(* IEC 61131-3 sources: daoli-st-library/DL_Process (part 66) *)

(* ---- FB_DL_InertPurgeSeq.st ---- *)
(*==============================================================================
 * 组件名称 (Component)  : FB_DL_InertPurgeSeq
 * 溯源说明 (Provenance): 道莅 clean-room 防御性实现（IEC 61131-3 纯净实现，闭源文档仅借语义，零代码行）
 * 所属子库 (Sublibrary) : DL_Process / Sequence
 * 当前版本 (Version)    : 1.0.0
 * 兼容性   (Platform)   : CODESYS 3.5 / TwinCAT 3 / 汇川 InoProShop / 施耐德
 *                         Machine Expert；纯 IEC 61131-3（第 3 版），仅用
 *                         Standard.library 的 TON / TIME_TO_DINT / DINT_TO_TIME
 * 组件分类 (Category)   : 功能块（FUNCTION_BLOCK）· 氮气置换顺控
 * 功能一句话 (Summary)  : 抽真空 → 充氮 → 保压取样 三相同循环置换，氧含量达目标
 *                         即放行，循环耗尽未达标则锁定失败，中止任意拍立即停。
 *
 * 本件存在的意义 (Why this unit exists)
 *   可燃溶剂场合点火/投料前的氮气置换是强制步骤，也是审核最容易被问的
 *   一条。它的逻辑不难，但「相转出必须断输入」这一点几乎每份手写代码都会
 *   踩：三相共用一只 TON，抽真空相残留的 ET 会让充氮相提前结束，或者
 *   保压相一进就走。本件把每相各一只 TON、相转出断输入一拍写成结构约束
 *   （R40 家族第三次事故的共同形态就在这一格）。
 *
 * 单循环定义 (One cycle)
 *   eEvacuate   : 抽真空阀开，tEvac 时间到**且**真空达 fVacOk → 进充氮
 *   eFillN2     : 充氮阀开，tFill 时间到 → 进保压取样
 *   eHoldVerify : 全阀关（保持压力），tHold 后读取氧含量
 *                 ≤ fO2Target → eComplete（信息 01DF）
 *                 否则循环数 +1：未达 uMaxCycles → eCycleDone → 回抽真空（信息 01DE）
 *                 已达 uMaxCycles → eFailed（故障 0313）
 *
 * 中止语义（三件顺控件共用同一段口径）
 *   bAbort **任意拍**生效：先清全部执行输出（三相阀），再回 eIdle；
 *   **不排队、不回退重来、不自动续跑**——中止是人的决定，重启必须由新的
 *   bStart 重新开始。原因：自动续跑会让操作工以为按了一次中止就断电了，
 *   实际设备又自己动起来，这是顺控件最危险的一类行为（R34 家族）。
 *
 * 边界安全 (Boundary)
 *   ① fO2Target <= 0、uMaxCycles = 0 或任一 TIME = 0 → 故障 0311、回 eIdle；
 *   ② bO2SensorOk = FALSE → 故障 0312、**禁止放行**（bDone 恒 FALSE）、三阀全关；
 *      氧分析仪坏掉时置换结果无从判断，继续循环只是白烧氮气；
 *   ③ 循环耗尽未达标 → bFailed := TRUE + 故障 0313；
 *   ④ 抽真空相 tEvac 到而真空未达 → 重新计时继续抽，连续 DL_EVAC_RETRY 次仍未达
 *      → 按「置换无法建立」处理，复用 0313（R90 不加码，理由见头注释）；
 *   ⑤ 三相各一只 TON，相转出以「断输入一拍」标志重启，绝不跨相复用实例；
 *   ⑥ 三阀输出互斥，段 1 先全清、段 7 按状态最多置一路（R72）；
 *   ⑦ CASE 落 ELSE 置 0313 并回 eIdle（兜底复用，R90）；
 *   ⑧ 放空阀编排约定：仅在 eComplete（置换合格）后打开以便泄压放行；
 *      eFailed 与其它相一律关闭——置换失败时保持惰化封闭，交人工处置。
 *
 * 引脚补全声明 (Pin completion)
 *   规格正文要求「真空达 fVacOk」判据，但引脚表未列真空度实测，故补
 *   fVacMeas : REAL [kPa g]。缺此引脚则「抽真空到位」无从判断，只能退化成
 *   纯定时，与本件语义不符。
 *
 * 错误码    : 16#0005_01DE 单循环未达标，进入下一循环——信息级
 *             16#0005_01DF 取样窗内氧含量已达目标——信息级，放行前置条件满足
 *             16#0005_0311 置换参数非法（目标/循环数/时长）——故障级，回 eIdle
 *             16#0005_0312 氧分析仪无效，禁止放行——故障级，三阀全关
 *             16#0005_0313 置换循环耗尽未达标（含状态机兜底与真空建立失败复用，R90）——故障级
 * 码位总账  : 16#0005_01DE 用 / 16#0005_01DF 用 ｜ 16#0005_0311 用 / 16#0005_0312 用 / 16#0005_0313 用
 * 状态机    : E_DL_PurgeState（eIdle / eEvacuate / eFillN2 / eHoldVerify / eCycleDone /
 *             eComplete / eFailed / eFault），CASE 含 ELSE 兜底，ELSE 置 16#0005_0313 并回 eIdle
 * 采样约定  : 每任务周期调用一次；各相时长由引脚给定，不读系统时钟
 * 依赖说明  : 只做组合编排，不复制低层算法；无 DL_ 子库调用
 * 验收向量  : V1 启动 → 抽真空 60 s 且真空 −85 kPa（< −80）→ 充氮 60 s → 保压 30 s
 *               读到 O2 1.2 %（≤ 2.0）→ eComplete，bDone = TRUE，eErr = 01DF
 *             V2 保压后 O2 3.5 %（> 2.0）、uMaxCycles = 3 → uCycleDone = 1，eErr = 01DE，
 *                回抽真空继续（循环主向量）
 *             V3 V2 连续三次未达标 → eFailed，bFailed = TRUE，eErr = 0313（耗尽主向量）
 *             V4 抽真空相 bAbort = TRUE → 三阀同拍全 FALSE，回 eIdle，不续跑（中止主向量）
 *             V5 bO2SensorOk = FALSE → eFault，三阀全关，bDone 恒 FALSE，eErr = 0312
 *             V6 uMaxCycles = 0 → eFault，eErr = 0311，回 eIdle
 *             V7 抽真空 3 次定时到但真空只有 −50 kPa → eFailed，eErr = 0313（真空建立失败复用）
 *             V8 eComplete 且 bStart 仍为 TRUE → 保持 eComplete（不放行丢失）；bStart 落 → eIdle
 * 红线自检  : 全局变量声明零使用 / 外部变量访问零使用 / 物理地址零使用 ｜ 纯 IEC 61131-3 ｜ 无除法
 *             浮点只用大小比较 ｜ 无循环 ｜ 全变量双语同行注释 ｜ ENUM + CASE 含 ELSE
 *             ｜ 三只 TON 在主体前部无条件刷新且各相各一只 ｜ 单拍标志全部预清零
 *             ｜ 阈值常量化，无魔法数
 * 修订历史  : 2026-11-16  v1.0.0  首版入库（R22 · 批 3 · 批处理顺控）
 *============================================================================*)

(*-----------------------------------------------------------------------------
 * 枚举: E_DL_PurgeState（归属本功能块，同文件发布，全库唯一定义）
 * 含义: 氮气置换顺控相位，每个成员在 CASE 中有且仅有一个标签。
 *-----------------------------------------------------------------------------*)
TYPE E_DL_PurgeState :
(
    eIdle       := 0,   // 待机：未启动或已复位 / Idle, not started or already reset
    eEvacuate   := 10,  // 抽真空相：真空阀开 / Evacuation, vacuum valve open
    eFillN2     := 20,  // 充氮相：氮气阀开 / Nitrogen fill, nitrogen valve open
    eHoldVerify := 30,  // 保压取样相：全阀关，读氧含量 / Hold and verify, all valves closed
    eCycleDone  := 40,  // 单循环结束（单拍相），随后回抽真空 / Cycle done, one scan then back to evacuation
    eComplete   := 50,  // 置换合格：放行 / Complete, production released
    eFailed     := 60,  // 置换失败锁定：循环耗尽 / Failed, cycles exhausted and latched
    eFault      := 99   // 故障：参数非法或氧分析仪无效 / Fault, illegal parameters or an invalid oxygen analyser
);
END_TYPE

FUNCTION_BLOCK FB_DL_InertPurgeSeq
VAR_INPUT
    bStart       : BOOL;                       // 启动请求，电平有效 / start request, level active
    bAbort       : BOOL;                       // 中止请求，任意拍生效 / abort request, effective on any scan
    fO2Meas      : REAL;                       // 氧含量实测 [%] / measured oxygen content [%]
    bO2SensorOk  : BOOL;                       // 氧分析仪有效性 / oxygen analyser validity
    fO2Target    : REAL := 2.0;                // 目标氧含量 [%]，须 > 0 / target oxygen content [%], must be > 0
    uMaxCycles   : UINT := 3;                  // 最大置换循环数 [次]，须 > 0 / maximum purge cycles [count], must be > 0
    tEvac        : TIME := T#60S;              // 抽真空时长 [ms]，须 > 0 / evacuation duration [ms], must be > 0
    tFill        : TIME := T#60S;              // 充氮时长 [ms]，须 > 0 / nitrogen fill duration [ms], must be > 0
    tHold        : TIME := T#30S;              // 保压取样时长 [ms]，须 > 0 / hold and verify duration [ms], must be > 0
    fVacOk       : REAL := -80.0;              // 抽真空到位阈值 [kPa g]，读数须 <= 本值 / vacuum target [kPa g]
    fVacMeas     : REAL;                       // 真空度实测 [kPa g]（引脚补充，见头注释） / measured vacuum [kPa g]
END_VAR
VAR_OUTPUT
    bVacValveCmd  : BOOL;                      // 抽真空阀指令 / vacuum valve command
    bN2ValveCmd   : BOOL;                      // 氮气阀指令 / nitrogen valve command
    bVentValveCmd : BOOL;                      // 放空阀指令（仅合格后打开） / vent valve command, opened only when qualified
    uCycleDone    : UINT;                      // 已完成置换循环数 [次] / completed purge cycles [count]
    bDone         : BOOL;                      // 置换合格放行 / purge qualified, production released
    bFailed       : BOOL;                      // 置换失败锁定 / purge failed, latched
    eErr          : UDINT;                     // 错误码，0 表示无错 / error code, 0 means no error
    bError        : BOOL;                      // 故障级标志，仅故障级错误置位 / fault-class flag, set only on fault-level codes
    bValid        : BOOL;                      // 输出可用标志 / outputs usable flag
END_VAR
VAR
    fbEvac       : TON;                        // 抽真空相计时，段 5 无条件刷新 [ms] / evacuation timer
    fbFill       : TON;                        // 充氮相计时，段 5 无条件刷新 [ms] / nitrogen fill timer
    fbHold       : TON;                        // 保压取样相计时，段 5 无条件刷新 [ms] / hold and verify timer
    _eState      : E_DL_PurgeState := E_DL_PurgeState.eIdle; // 当前相位 / current phase
    _bInit       : BOOL := FALSE;              // 首扫标志，初值 FALSE 取非判定 / first-scan flag, tested negated
    _bParamBad   : BOOL;                       // 参数非法标志 / illegal parameter flag
    _bSensorBad  : BOOL;                       // 氧分析仪无效标志 / invalid analyser flag
    _bIllegal    : BOOL;                       // 非法状态标志 / illegal state flag
    _bEvacBreak  : BOOL;                       // 抽真空计时器断输入一拍 / evacuation timer one-scan break
    _bFillBreak  : BOOL;                       // 充氮计时器断输入一拍 / fill timer one-scan break
    _bHoldBreak  : BOOL;                       // 保压计时器断输入一拍 / hold timer one-scan break
    _bVacOk      : BOOL;                       // 真空到位判据 / vacuum reached
    _bQualified  : BOOL;                       // 本拍取样合格 / qualified this scan
    _bCycleEvent : BOOL;                       // 本拍单循环结束事件 / cycle finished this scan
    _uCycleAcc   : UINT;                       // 已完成循环数保持量 [次] / held completed cycle count
    _uEvacRetry  : UINT;                       // 抽真空重试计数 [次] / evacuation retry counter
    _bFailedAcc  : BOOL;                       // 失败锁存保持量 / held failure latch
END_VAR
VAR CONSTANT
    DL_VAL_LIM     : REAL := 1.0E6;            // 有限性判定的绝对值上限 [无量纲] / finiteness ceiling
    DL_O2_MIN      : REAL := 0.0;              // 目标氧含量下限 [%]，须严格大于 / target oxygen floor, strictly greater
    DL_CYCLE_MIN   : UINT := 0;                // 循环数下限 [次] / cycle floor [count]
    DL_EVAC_RETRY  : UINT := 3;                // 抽真空最大重试次数 [次] / maximum evacuation retries
    DL_TIME_ZERO   : TIME := T#0MS;            // 时间零值基准 [ms] / time zero reference
    DL_CNT_MAX     : UINT := 65535;            // 循环计数饱和上界 [次] / cycle count saturation ceiling
END_VAR

(*------------------------------------------------------------------------------
 * 段 1｜每拍预置：三阀**先全清**（R72），单拍标志预清零（R25 第一律）
 *      Both commands cleared first, one-shot flags pre-cleared
 *-----------------------------------------------------------------------------*)
bVacValveCmd  := FALSE;                        // 抽真空阀先清 / vacuum valve cleared first
bN2ValveCmd   := FALSE;                        // 氮气阀先清 / nitrogen valve cleared first
bVentValveCmd := FALSE;                        // 放空阀先清 / vent valve cleared first
bDone         := FALSE;                        // 放行标志每拍重算 / release flag recomputed
bFailed       := FALSE;                        // 失败标志每拍重算 / failure flag recomputed
bValid        := FALSE;                        // 可用标志每拍重算 / usable flag recomputed
eErr          := 16#0000_0000;                 // 错误码每拍重算 / error code recomputed
bError        := FALSE;                        // 故障标志每拍重算 / fault flag recomputed
_bParamBad    := FALSE;                        // 参数非法标志预清零 / parameter flag pre-cleared
_bSensorBad   := FALSE;                        // 分析仪无效标志预清零 / analyser flag pre-cleared
_bIllegal     := FALSE;                        // 非法状态标志预清零 / illegal state flag pre-cleared
_bVacOk       := FALSE;                        // 真空到位判据预置 FALSE / vacuum reached preset FALSE
_bQualified   := FALSE;                        // 合格判据预置 FALSE / qualified preset FALSE
_bCycleEvent  := FALSE;                        // 循环事件预置 FALSE / cycle event preset FALSE

(*------------------------------------------------------------------------------
 * 段 2｜首扫初始化（循环计数与失败锁存从零起）
 *      First-scan initialisation
 *-----------------------------------------------------------------------------*)
IF NOT _bInit THEN
    _eState      := E_DL_PurgeState.eIdle;     // 相位待机 / phase idle
    _uCycleAcc   := 0;                         // 循环计数清零 [次] / cycle count cleared
    _uEvacRetry  := 0;                         // 重试计数清零 [次] / retry counter cleared
    _bFailedAcc  := FALSE;                     // 失败锁存清零 / failure latch cleared
    _bEvacBreak  := TRUE;                      // 抽真空计时从零开始 / evacuation timer starts from zero
    _bFillBreak  := TRUE;                      // 充氮计时从零开始 / fill timer starts from zero
    _bHoldBreak  := TRUE;                      // 保压计时从零开始 / hold timer starts from zero
    _bInit       := TRUE;                      // 首扫只做一次 / the first scan runs once
END_IF

(*------------------------------------------------------------------------------
 * 段 3｜参数闸门（目标氧含量、循环数、三相时长）
 *      Parameter gate for the target, the cycle count and the three durations
 *-----------------------------------------------------------------------------*)
IF (fO2Target <> fO2Target) OR (ABS(fO2Target) > DL_VAL_LIM) OR (fO2Target <= DL_O2_MIN) THEN
    _bParamBad := TRUE;                        // 目标氧含量非法 / target oxygen illegal
END_IF
IF uMaxCycles <= DL_CYCLE_MIN THEN
    _bParamBad := TRUE;                        // 循环数为 0，置换无从进行 / zero cycles, nothing to run
END_IF
IF (TIME_TO_DINT(tEvac) <= 0) OR (TIME_TO_DINT(tFill) <= 0) OR (TIME_TO_DINT(tHold) <= 0) THEN
    _bParamBad := TRUE;                        // 任一相时长为 0 / a phase duration is zero
END_IF

(*------------------------------------------------------------------------------
 * 段 4｜氧分析仪有效性与真空判据（分析仪坏掉时禁止放行）
 *      Analyser validity and the vacuum test
 *-----------------------------------------------------------------------------*)
IF NOT bO2SensorOk THEN
    _bSensorBad := TRUE;                       // 分析仪无效 / the analyser is invalid
END_IF
_bVacOk := (fVacMeas <= fVacOk);               // 真空到位：读数不高于阈值（越负越真空） / reached when the reading is deep enough

(*------------------------------------------------------------------------------
 * 段 5｜三只计时器无条件刷新（R40：CASE 之外每拍必调；**一相一只，绝不共用**）
 *      Three timers refreshed unconditionally, one per phase, never shared
 *-----------------------------------------------------------------------------*)
fbEvac(IN := (_eState = E_DL_PurgeState.eEvacuate) AND (NOT _bEvacBreak), PT := tEvac); // 抽真空相计时
_bEvacBreak := FALSE;                          // 断输入拍在调用后自清 / break self-cleared after the call

fbFill(IN := (_eState = E_DL_PurgeState.eFillN2) AND (NOT _bFillBreak), PT := tFill); // 充氮相计时
_bFillBreak := FALSE;                          // 断输入拍在调用后自清 / break self-cleared after the call

fbHold(IN := (_eState = E_DL_PurgeState.eHoldVerify) AND (NOT _bHoldBreak), PT := tHold); // 保压取样相计时
_bHoldBreak := FALSE;                          // 断输入拍在调用后自清 / break self-cleared after the call

(*------------------------------------------------------------------------------
 * 段 6｜相位机（只做迁移；阀输出在段 7）
 *      Phase machine, transitions only, the valve commands are set in segment seven
 *-----------------------------------------------------------------------------*)
IF bAbort THEN
    (* 中止：任意拍生效，先清输出（段 1 已清）再回待机，不排队不回退 *)
    (* Abort takes effect on any scan, no queuing and no rollback *)
    _eState     := E_DL_PurgeState.eIdle;
    _uEvacRetry := 0;                          // 重试计数清零 [次] / retry counter cleared
    _bEvacBreak := TRUE;                       // 三相计时全部重启 / every timer restarts
    _bFillBreak := TRUE;
    _bHoldBreak := TRUE;
ELSIF _bParamBad THEN
    _eState := E_DL_PurgeState.eFault;         // 参数非法：转故障 / illegal parameters go to fault
    _bEvacBreak := TRUE;                       // 计时重启，避免把故障期算进相时长 / timers restart
    _bFillBreak := TRUE;
    _bHoldBreak := TRUE;
ELSIF _bSensorBad THEN
    _eState := E_DL_PurgeState.eFault;         // 分析仪无效：转故障，三阀全关（段 7 自然全关） / invalid analyser
    _bEvacBreak := TRUE;                       // 计时重启 / timers restart
    _bFillBreak := TRUE;
    _bHoldBreak := TRUE;
ELSE
    CASE _eState OF

        E_DL_PurgeState.eIdle:                 // 待机：启动即从第一个循环开始
            IF bStart THEN
                _uCycleAcc  := 0;              // 新任务循环数从零起 [次] / a new job starts at zero cycles
                _uEvacRetry := 0;              // 重试计数清零 [次] / retry counter cleared
                _bFailedAcc := FALSE;          // 失败锁存清零 / failure latch cleared
                _bEvacBreak := TRUE;           // 抽真空计时从零开始 / the evacuation timer starts from zero
                _eState     := E_DL_PurgeState.eEvacuate; // 进抽真空相 / enter evacuation
            END_IF

        E_DL_PurgeState.eEvacuate:             // 抽真空：时间到且真空到位才转充氮
            IF NOT bStart THEN
                _eState := E_DL_PurgeState.eIdle; // 启动撤销，回待机（等价于中止） / start dropped
            ELSIF fbEvac.Q AND _bVacOk THEN
                _uEvacRetry := 0;              // 本次抽真空成功，重试计数清零 / evacuation succeeded
                _bFillBreak := TRUE;           // 充氮计时从零开始（相转出断输入） / the fill timer starts from zero
                _eState     := E_DL_PurgeState.eFillN2; // 进充氮相 / enter the fill phase
            ELSIF fbEvac.Q THEN
                _uEvacRetry := _uEvacRetry + 1; // 时间到但真空未达：重试累计 / elapsed without vacuum, retry counted
                _bEvacBreak := TRUE;           // 抽真空计时重启 / the evacuation timer restarts
                IF _uEvacRetry >= DL_EVAC_RETRY THEN
                    _bFailedAcc := TRUE;       // 真空建立失败：按失败锁定处理 / the vacuum cannot be established
                    _eState     := E_DL_PurgeState.eFailed;
                END_IF
            END_IF

        E_DL_PurgeState.eFillN2:               // 充氮：时间到即转保压取样
            IF NOT bStart THEN
                _eState := E_DL_PurgeState.eIdle; // 启动撤销，回待机 / start dropped
            ELSIF fbFill.Q THEN
                _bHoldBreak := TRUE;           // 保压计时从零开始（相转出断输入） / the hold timer starts from zero
                _eState     := E_DL_PurgeState.eHoldVerify; // 进保压取样相 / enter hold and verify
            END_IF

        E_DL_PurgeState.eHoldVerify:           // 保压取样：窗满读氧含量
            IF NOT bStart THEN
                _eState := E_DL_PurgeState.eIdle; // 启动撤销，回待机 / start dropped
            ELSIF fbHold.Q THEN
                _bCycleEvent := TRUE;          // 单循环结束事件（段 7 消费） / the cycle finished
            END_IF

        E_DL_PurgeState.eCycleDone:            // 单循环结束（单拍相）：回抽真空
            _bEvacBreak := TRUE;               // 抽真空计时从零开始（相转出断输入） / the evacuation timer restarts
            _uEvacRetry := 0;                  // 重试计数按循环清零 [次] / retries reset per cycle
            _eState     := E_DL_PurgeState.eEvacuate; // 进下一循环 / next cycle
        E_DL_PurgeState.eComplete:             // 合格：等启动撤销才可复位
            IF NOT bStart THEN
                _eState := E_DL_PurgeState.eIdle; // 启动撤销，回待机 / back to idle once the start drops
            END_IF

        E_DL_PurgeState.eFailed:               // 失败锁定：等启动撤销才可复位
            IF NOT bStart THEN
                _eState := E_DL_PurgeState.eIdle; // 启动撤销，回待机 / back to idle once the start drops
            END_IF

        E_DL_PurgeState.eFault:                // 故障：参数与分析仪恢复且未启动才回待机
            IF (NOT _bParamBad) AND (NOT _bSensorBad) AND (NOT bStart) THEN
                _eState := E_DL_PurgeState.eIdle; // 原因消失 / the cause is gone
            END_IF

        ELSE
            _bIllegal := TRUE;                 // 标记非法状态 / flag the illegal state
            _bEvacBreak := TRUE;               // 三相计时重启 / every timer restarts
            _bFillBreak := TRUE;
            _bHoldBreak := TRUE;
            _eState := E_DL_PurgeState.eIdle;  // 回安全态 / back to the safe state
        END_CASE
END_IF

(*------------------------------------------------------------------------------
 * 段 7｜单循环判定与阀输出（互斥：段 1 已全清，此处最多置一路）
 *      Cycle verdict and valve commands, at most one is set here
 *-----------------------------------------------------------------------------*)
IF _bCycleEvent THEN
    _bQualified := (fO2Meas <= fO2Target);     // 氧含量达目标即合格 [布尔] / qualified when the oxygen reaches the target
    IF _bQualified THEN
        _eState := E_DL_PurgeState.eComplete;  // 合格：放行 / qualified, release
    ELSE
        IF _uCycleAcc < DL_CNT_MAX THEN
            _uCycleAcc := _uCycleAcc + 1;      // 循环数 +1（饱和不回绕） [次] / cycle count incremented
        END_IF
        IF _uCycleAcc >= uMaxCycles THEN
            _bFailedAcc := TRUE;               // 循环耗尽：失败锁定 / cycles exhausted, latch the failure
            _eState     := E_DL_PurgeState.eFailed;
        ELSE
            _eState := E_DL_PurgeState.eCycleDone; // 进下一循环 / next cycle
        END_IF
    END_IF
    _bHoldBreak := TRUE;                       // 离开保压相，计时重启 / leave hold, restart the timer
END_IF

CASE _eState OF
    E_DL_PurgeState.eEvacuate:                 // 抽真空阀开 / vacuum valve open
        bVacValveCmd := TRUE;
    E_DL_PurgeState.eFillN2:                   // 氮气阀开 / nitrogen valve open
        bN2ValveCmd := TRUE;
    E_DL_PurgeState.eComplete:                 // 合格后放空泄压放行 / vent only when qualified
        bVentValveCmd := TRUE;
    ELSE
        bVacValveCmd  := FALSE;                // 其余相：显式重申全关（R72 双路径） / explicitly re-asserted closed
        bN2ValveCmd   := FALSE;
        bVentValveCmd := FALSE;
END_CASE

(*------------------------------------------------------------------------------
 * 段 8｜码位优先级链与出口
 *      Code priority chain and exit
 *-----------------------------------------------------------------------------*)
IF _bIllegal THEN
    _bFailedAcc := TRUE;                       // 非法状态按失败锁定处理 / an illegal state latches a failure
END_IF

IF _bParamBad THEN
    eErr   := 16#0005_0311;                    // 故障级：置换参数非法 / fault: purge parameters illegal
    bError := TRUE;                            // 置故障标志 / raise the fault flag
    _eState := E_DL_PurgeState.eIdle;          // 明确回待机（参数非法不谈顺控） / back to idle
ELSIF _bSensorBad THEN
    eErr   := 16#0005_0312;                    // 故障级：氧分析仪无效，禁止放行 / fault: analyser invalid, release forbidden
    bError := TRUE;                            // 置故障标志 / raise the fault flag
    bVacValveCmd  := FALSE;                    // 三阀显式全关（禁止放行的实际动作） / all valves explicitly closed
    bN2ValveCmd   := FALSE;
    bVentValveCmd := FALSE;
ELSIF (_eState = E_DL_PurgeState.eFailed) OR _bFailedAcc THEN
    eErr   := 16#0005_0313;                    // 故障级：循环耗尽未达标（兜底与真空失败复用） / fault: cycles exhausted
    bError := TRUE;                            // 置故障标志 / raise the fault flag
ELSIF _bIllegal THEN
    eErr   := 16#0005_0313;                    // 故障级：非法状态兜底（同一码，R90） / fault: illegal state fallback
    bError := TRUE;                            // 置故障标志 / raise the fault flag
ELSIF _eState = E_DL_PurgeState.eComplete THEN
    eErr   := 16#0005_01DF;                    // 信息级：取样窗内氧含量已达目标 / informational: the target was reached
ELSIF _bCycleEvent THEN
    eErr   := 16#0005_01DE;                    // 信息级：单循环未达标，进入下一循环 / informational: next cycle
END_IF

uCycleDone := _uCycleAcc;                      // 已完成循环数出口 [次] / completed cycles outlet
bDone      := (_eState = E_DL_PurgeState.eComplete); // 放行出口：仅合格相为真 / release outlet
bFailed    := (_eState = E_DL_PurgeState.eFailed) OR _bFailedAcc; // 失败出口 / failure outlet

IF bError OR _bSensorBad THEN
    bValid := FALSE;                           // 故障级或分析仪无效：输出不可用 / fault or invalid analyser: unusable
ELSIF _bParamBad THEN
    bValid := FALSE;                           // 参数非法：输出不可用 / illegal parameters: unusable
ELSE
    bValid := TRUE;                            // 输出可用（顺控进行中亦可用） / usable, also while running
END_IF

END_FUNCTION_BLOCK

(* ---- FB_DL_LeakTestStation.st ---- *)
(*==============================================================================
 * 组件名称 (Component)  : FB_DL_LeakTestStation
 * 所属子库 (Sublibrary) : DL_Process
 * 当前版本 (Version)    : 1.0.2
 * 兼容性 (Platform)   : CODESYS 3.5 / TwinCAT 3 / 汇川 InoProShop / Machine Expert
 *                         仅依赖 Standard.library（TON / R_TRIG），零厂商方言
 * 分类     (Category)   : 工艺段功能块（Function Block · 压降法气密检漏工站）
 * 功能简述 (Function)   : 压降法气密检漏十相顺控：夹具确认 → 充气 → 稳压 →
 *                         隔离测量 → 排气 → PASS/NG/Abort。内置大漏快判、温
 *                         度补偿（一阶理想气体近似）、稳压超容差设备异常与工
 *                         件不良分离判定（工件 NG 不置故障位）。本工站为流程
 *                         编排与判定层——检漏仪精度与夹具密封属测量系统，不
 *                         在本块职责内；压力/温度反馈由调用方适配层注入。
 * 首扫说明 (Init note)  : 顺序型组件但全部状态由指令沿/电平驱动，无跟踪/初
 *                         始化语义，免首扫（R23/公约 0.1），无 bInit。
 * 公约遵循 (Convention) : 0.2/R21 bError 仅故障级码置位（工件 NG 不置位）；
 *                         0.4 双语同行注释；0.5/R7 实例主体最前部无条件刷新；
 *                         0.10 定时基准由引脚给——依公约增补 tCycle 输入引
 *                         脚（泳道 A FB_DL_ElectronicGear 同款处理，公共约
 *                         定强制项，非逐组件条款）；0.14 非有限值自比等价式
 *                         防御、除法前判零；0.15 压力统一 kPa、温度统一 ℃、
 *                         泄漏率统一 mL/min，同块不混用同类单位；0.16 无魔
 *                         法数；0.17 终结符成对 ✓；0.19 码位同行【级别】注
 *                         释；0.20 验收向量入头注释；R25 bDone 单拍三律；
 *                         R14 语义参数（各相计时 PT）变更经相位切换自然断输
 *                         入一拍归零。
 * 红线自检 (Redline)    : R1 零全局变量表/外部变量引用 ✓｜R2 零物理 IO 地址 ✓
 *                         R3 纯 IEC 61131-3 ✓｜R4 非有限值/除零/互斥出口 ✓
 *                         R5 全变量中英双语同行注释 ✓｜R6 ENUM+CASE+ELSE ✓
 *                         R7 七实例（R_TRIG×2/TON×5）主体最前部无条件刷新 ✓
 *                         R8 全常量化 ✓｜R25 单拍标志生命周期三律 ✓
 * 设计要点 (Key notes)  : ① 充气出口双条件：最小充气保持时长 tFill 到且压力
 *                           达 target×(1−DL_LEAK_FILL_TOL)——tFill 按「最小
 *                           充气保持时长」实现（偏离留档②）；
 *                         ② 稳压结束压力超容差 → 故障 0252 设备异常（不判工
 *                           件 NG，测量系统与被测件责任分离）；
 *                         ③ 大漏快判：测量窗内压降 ≥ fGrossLeakDrop 立即 NG
 *                           （信息码 0153），fGrossLeakDrop=0 禁用快判；
 *                         ④ 泄漏率量纲推导（完整链）：Q[kPa·mL/s] = ΔP[kPa]
 *                           × V[mL] / t[s]；乘 DL_LEAK_UNIT_FACTOR=60 转分钟
 *                           口径 → Q[mL/min]。该系数为工艺约定换算（秒→分），
 *                           非严格气体动力学模型；温度补偿
 *                           Q ×= (273.15+fRefTemp)/(273.15+fT0) 为一阶理想气
 *                           体近似，适用于温漂小、测量窗短的常规检漏工况；
 *                         ⑤ 压差回负（温度回升）按 0 处理 + 信息码 0151，不
 *                           判 NG；bPass/bFail 先清后置保证互斥出口；
 *                         ⑥ 秒值换算：测量时长经 tCycle 引脚折算（TIME 毫
 *                           秒口径 /1000，TIME_TO_REAL），tCycle 非有限值/
 *                           非正 → 故障 0254 归并（输入防御）。
 * 偏离留档 (Deviation)  : 依 R11 头注释留档，共 2 条：
 *                         ① tCycle 增补引脚：规格引脚表未含任务周期，泄漏率
 *                           秒值换算必须有时间基准；理由/影响见公约 0.10 与
 *                           泳道 A 先例——公共约定强制项，非语义偏离；
 *                         ② tFill 引脚语义展开：规格仅列「充气时长」未定义
 *                           出口关系，按「最小充气保持时长（到时才允许判压
 *                           力达标）」实现；理由：防止大容积腔体压力冲击期误
 *                           判达标；影响：充气相出口 = tFill 到 AND 压力达标
 *                           双条件，仅接压力反馈而不接 tFill 的调用方需给足
 *                           tFill=最小值。
 * 开源溯源 (Origin)     : 来源标签 leak-test / pressure-decay（RAW_NOTES_R8
 *                         S-8：压降法检漏公开工程惯例——充气/稳压/隔离测量/
 *                         排气相序、测量前必须隔离气源、稳压过短既藏漏又造
 *                         漏、大漏表现为充不上压、稳压超容差属设备异常（提取
 *                         点⑤⑥），公开技术资料，仅借鉴相序分类与参数域；状态
 *                         机、码位、引脚契约、温度补偿与量纲推导 100% 本库独
 *                         立设计，clean-room 未复制源码。许可证说明：借鉴对象
 *                         为公开技术惯例，无附带许可限制；本文件为本库原创实
 *                         现，随本库许可证发布）。
 * 验收向量 (Acceptance) :
 *   V1 合格件（ΔP 对应 Q < 限值）→ ePass + bDone 单拍 + nPartCount +1；
 *   V2 大漏件（充不上压）→ 充气超时 0251；
 *   V3 测量窗 ΔP 超快判阈 → 立即 FAIL + 信息码 0153；
 *   V4 稳压结束压力超容差 → 0252 且不判 NG（设备异常分离）；
 *   V5 温度 35 ℃ 时补偿后 Q 下降（比值 298.15/308.15）；
 *   V6 bAbort 测量中 → 立即排气不记 NG、判定输出清；
 *   V7 fChamberVolume=0 → 0255（除零防护）；
 *   V8 排气超时 → 0253。
 * 修订历史 (Revision)   :
 *   2026-11-15  v1.0.0  首版入库（Round 08 · DL_Process 检漏工站件）
 *   2026-11-15  v1.0.1  R8 总监终审修复：终端态分支内的孤立空语句 `;`（非 IEC 61131-3 文法，statement_list 允许零条语句但不容纳孤立分号）改为纯注释占位分支，行为等价、跨平台可移植性合规。
 *   2026-11-15  v1.0.2  R11 修复：压差锁存赋值目标笔误，`_fDeltaP` -> `fDeltaP`（输出 fDeltaP 此前全文零写入致恒 0，属功能缺口 + 未声明标识符编译阻断双缺陷）；快判路径与测量结算路径各一处，共 2 处。
 *                       R11 fix: assignment target erratum, `_fDeltaP` -> `fDeltaP` (2 sites).
 *============================================================================*)

(*-----------------------------------------------------------------------------
 * 枚举: E_DL_LeakPhase（归属 FB_DL_LeakTestStation，与其同文件发布，公约 0.18）
 *----------------------------------------------------------------------------*)
TYPE E_DL_LeakPhase :
(
    eIdle       := 0,   // 空闲：等启动 / Idle, awaiting start
    eClampCheck := 10,  // 夹具确认：等夹具闭合信号 / Clamp check, awaiting fixture closed
    eFill       := 20,  // 充气：充气阀开，至目标压力 / Fill, valve open to target pressure
    eStabilize  := 30,  // 稳压：隔离保温，等热平衡 / Stabilize, isolated for thermal balance
    eMeasure    := 40,  // 测量：隔离测压降 / Measure, isolated pressure-decay window
    eVent       := 50,  // 排气：排气阀开，泄压到安全位 / Vent, depressurize to safe level
    ePass       := 60,  // 合格：结果保持，等复位/新周期 / Pass verdict held
    eFail       := 70,  // 不合格：结果保持，等复位 / Fail verdict held
    eAbort      := 80,  // 中止：操作员/上游中止，安全排气 / Aborted, safe depressurize
    eFault      := 99   // 设备故障锁存 / Equipment fault latched
) UINT;
END_TYPE

FUNCTION_BLOCK FB_DL_LeakTestStation
VAR_INPUT
    bEnable             : BOOL;             // 工站使能（Station enable），FALSE=安全排气并清判定输出 / Enable, FALSE = safe depressurize and clear verdicts
    bStart              : BOOL;             // 启动测试周期（Start），上升沿受理（空闲/合格/不合格态）/ Start edge accepted at idle/pass/fail
    bAbort              : BOOL;             // 中止（Abort），电平最高优先 → 安全排气 / Abort level, highest priority, safe vent
    bReset              : BOOL;             // 复位故障与结果（Reset），上升沿受理 / Rising edge resets fault and verdicts
    bFixtureClosed      : BOOL;             // 夹具闭合确认（Fixture closed），FALSE 禁止充气 / Fixture closed interlock, FALSE blocks fill
    bTempCompEnable     : BOOL := TRUE;     // 温度补偿使能（Temp compensation），FALSE=按原始压降计算 / Temperature compensation enable
    fTestPressure       : REAL := 300.0;    // 目标测试压力（Test pressure）[kPa]，域 1..10000 / Target test pressure [kPa]
    fPressureTol        : REAL := 5.0;      // 稳压结束压力容差（Pressure tolerance）[kPa]，域 0.1..100；超容差判设备异常 / Pressure tolerance at stabilize end [kPa]
    fActPressure        : REAL;             // 实际压力（Actual pressure）[kPa]，由变送器/适配层注入 / Actual pressure [kPa] injected by adapter
    fActTemp            : REAL := 25.0;     // 实际温度（Actual temperature）[℃]，温度补偿用 / Actual temperature [degC]
    fRefTemp            : REAL := 25.0;     // 基准温度（Reference temperature）[℃]，补偿基准 / Reference temperature [degC]
    fChamberVolume      : REAL := 100.0;    // 被测腔容积（Chamber volume）[mL]，泄漏率换算用 / Chamber volume [mL] for leak-rate conversion
    fLeakLimit          : REAL := 10.0;     // 泄漏率上限（Leak rate limit）[mL/min]，≤ 此值为 PASS / Leak rate limit [mL/min], PASS below
    fGrossLeakDrop      : REAL := 20.0;     // 大漏快判压降（Gross leak drop）[kPa]，测量窗内超此值立即 NG；0=禁用快判 / Gross-leak quick-judge drop [kPa], 0 disables
    tFill               : TIME := T#3S;     // 最小充气保持时长（Min fill hold，偏离留档②），到时才允许判压力达标 / Minimum fill hold time before pressure verdict
    tStabilize          : TIME := T#5S;     // 稳压时长（Stabilize time），过短既藏漏又造漏 / Stabilize time
    tMeasure            : TIME := T#10S;    // 测量时长（Measure time），T#0S 判故障 / Measure window duration
    tFillTimeout        : TIME := T#20S;    // 充气超时（Fill timeout），兼作夹具确认超时 / Fill timeout, also clamp-check timeout
    tVentTimeout        : TIME := T#10S;    // 排气超时（Vent timeout）/ Vent timeout
    tCycle              : TIME := T#10MS;   // 任务扫描周期（Task cycle time）[ms]，由调用方按实际任务给，泄漏率秒值换算基准（公约 0.10）/ Task cycle time, seconds conversion base
END_VAR
VAR_OUTPUT
    bCmdFillValve       : BOOL;             // 充气阀指令（Fill valve）/ Fill valve command
    bCmdIsolateValve    : BOOL;             // 隔离阀指令（Isolate valve），测量期间为 TRUE（测量前必须隔离气源）/ Isolate valve, TRUE during stabilize/measure
    bCmdVentValve       : BOOL;             // 排气阀指令（Vent valve）/ Vent valve command
    ePhase              : E_DL_LeakPhase := E_DL_LeakPhase.eIdle; // 当前相位（Current phase）/ Current phase
    bBusy               : BOOL;             // 周期执行中（Busy），夹具确认至排气态为 TRUE / TRUE from clamp check to vent
    bDone               : BOOL;             // 周期结束单拍脉冲（Done pulse），单拍生命周期三律 / One-scan verdict pulse
    bPass               : BOOL;             // 判定合格（PASS），合格保持态为 TRUE / PASS verdict held
    bFail               : BOOL;             // 判定不合格（FAIL），不合格保持态为 TRUE / FAIL verdict held
    fLeakRate           : REAL;             // 计算泄漏率（Leak rate）[mL/min]，已含温度补偿，测量后锁存 / Leak rate [mL/min] latched after measure
    fDeltaP             : REAL;             // 测量窗压降（Pressure drop）[kPa]，锁存 / Pressure drop [kPa] latched
    bError              : BOOL;             // 设备故障锁存（Error），仅故障级码；工件 NG 不置此位 / Equipment fault, fault codes only, part NG excluded
    uErrorId            : UDINT;            // 故障码（Error code），16#0005_xxxx 段，0=无故障 / Error code, fault-level priority
    nPartCount          : UDINT;            // 测试件数（Part counter），每次判定 +1 / Tested part counter
    nRejectCount        : UDINT;            // 不合格件数（Reject counter）/ Rejected part counter
END_VAR
VAR
    _ePhase             : E_DL_LeakPhase := E_DL_LeakPhase.eIdle; // 内部相位（Internal phase）/ Internal phase
    _bFaultLatch        : BOOL;             // 设备故障锁存标志（Fault latch flag），仅复位路径清除 / Fault latch, cleared only via reset path
    _uErrorIdInt        : UDINT;            // 内部故障级码寄存（Internal fault-level register）/ Internal fault-level register
    _uInfoCode          : UDINT;            // 本拍信息级码（Info code this cycle），瞬时型每拍重算 / Transient info code
    _bAbortActive       : BOOL;             // 中止激活（Abort active），电平锁存至排气完成 / Abort latched until vent completes
    _bPassLatched       : BOOL;             // 判定锁存（Verdict latch），TRUE=合格 / Verdict latch, TRUE = pass
    _bVerdictValid      : BOOL;             // 判定有效（Verdict valid），有已结算结果 / A settled verdict exists
    _fDtS               : REAL;             // 扫描周期秒值（Cycle time seconds）[s]，tCycle 折算 / Cycle time in seconds
    _fTestPressEff      : REAL;             // 生效目标压力（Effective test pressure）[kPa]，防御后值 / Sanitized test pressure
    _fTolEff            : REAL;             // 生效容差（Effective tolerance）[kPa] / Sanitized tolerance
    _fVolEff            : REAL;             // 生效容积（Effective volume）[mL] / Sanitized volume
    _fLeakLimEff        : REAL;             // 生效泄漏率上限（Effective leak limit）[mL/min] / Sanitized leak limit
    _fGrossEff          : REAL;             // 生效大漏阈（Effective gross-leak threshold）[kPa] / Sanitized gross-leak threshold
    _fP0                : REAL;             // 测量起点压力（Pressure at measure start）[kPa] / Pressure at measure start
    _fT0                : REAL;             // 测量起点温度（Temperature at measure start）[℃] / Temperature at measure start
    _fDeltaPInt         : REAL;             // 内部压差（Internal delta-P）[kPa]，回负按 0 / Internal delta-P, negative floored to zero
    _fMeasSec           : REAL;             // 测量累计秒值（Accumulated measure seconds）[s] / Accumulated measure seconds
    _fLeakRateInt       : REAL;             // 内部泄漏率（Internal leak rate）[mL/min] / Internal leak rate
    _fDenK              : REAL;             // 温度补偿分母（Compensation denominator）[K] / Compensation denominator in kelvin
    _fbTrigStart        : R_TRIG;           // 启动沿（Start edge detector）/ Start edge detector
    _fbTrigReset        : R_TRIG;           // 复位沿（Reset edge detector）/ Reset edge detector
    _fbTonClampTo       : TON;              // 夹具确认超时（Clamp-check timeout）/ Clamp-check timeout
    _fbTonFillMin       : TON;              // 最小充气保持（Min fill hold）/ Minimum fill hold
    _fbTonFillTo        : TON;              // 充气超时（Fill timeout）/ Fill timeout
    _fbTonStab          : TON;              // 稳压时长（Stabilize duration）/ Stabilize duration
    _fbTonMeas          : TON;              // 测量时长（Measure duration）/ Measure duration
    _fbTonVentTo        : TON;              // 排气超时（Vent timeout）/ Vent timeout
END_VAR
VAR CONSTANT
    DL_LEAK_REAL_MAX    : REAL := 3.4E38;   // 单精度有限值判据幅值（Finite magnitude bound）/ Finite magnitude bound for REAL inputs
    DL_LEAK_EPS         : REAL := 1.0E-6;   // 浮点防零容差（Float divide-guard epsilon）/ Float divide-guard epsilon
    DL_LEAK_FILL_TOL    : REAL := 0.02;     // 充气达标相对容差（Fill reach tolerance）[-]，目标压力的 2% / Fill reach tolerance fraction of target
    DL_LEAK_UNIT_FACTOR : REAL := 60.0;     // 泄漏率秒→分换算系数（Seconds-to-minutes factor）[-]，工艺约定换算 / Unit conversion factor, convention
    DL_LEAK_VENT_DONE   : REAL := 2.0;      // 排气完成压力（Vent-done pressure）[kPa]，低于此值视为安全 / Vent-done pressure threshold [kPa]
    DL_LEAK_KELVIN      : REAL := 273.15;   // 摄氏→开氏偏移（Celsius-to-kelvin offset）[K] / Celsius-to-kelvin offset
    DL_LEAK_PRESS_MIN   : REAL := 1.0;      // 目标压力域下限（Test pressure lower clamp）[kPa] / Test pressure lower clamp
    DL_LEAK_PRESS_MAX   : REAL := 10000.0;  // 目标压力域上限（Test pressure upper clamp）[kPa] / Test pressure upper clamp
    DL_LEAK_TOL_MIN     : REAL := 0.1;      // 容差域下限（Tolerance lower clamp）[kPa] / Tolerance lower clamp
    DL_LEAK_TOL_MAX     : REAL := 100.0;    // 容差域上限（Tolerance upper clamp）[kPa] / Tolerance upper clamp
    DL_TIME_MS_SCALE    : REAL := 1000.0;   // 毫秒→秒换算（Milliseconds-to-seconds scale）[-] / Milliseconds-to-seconds scale
    DL_LEAK_ERR_CLAMP   : UDINT := 16#0005_0250; // 0005_0250 夹具闭合超时【故障级】/ Fixture closed timeout, fault level
    DL_LEAK_ERR_FILL    : UDINT := 16#0005_0251; // 0005_0251 充气超时未达压（大漏常见表现）【故障级】/ Fill timeout, gross leak typical, fault level
    DL_LEAK_ERR_STAB    : UDINT := 16#0005_0252; // 0005_0252 稳压结束压力超容差（设备异常）【故障级】/ Stabilize-end pressure out of tolerance, equipment fault
    DL_LEAK_ERR_VENT    : UDINT := 16#0005_0253; // 0005_0253 排气超时【故障级】/ Vent timeout, fault level
    DL_LEAK_ERR_NAN     : UDINT := 16#0005_0254; // 0005_0254 压力/温度/容积/阈值输入非有限值【故障级】/ Non-finite process input, fault level
    DL_LEAK_ERR_VOL     : UDINT := 16#0005_0255; // 0005_0255 腔容积非法（≤0，除零防护）【故障级】/ Invalid chamber volume, fault level
    DL_LEAK_ERR_MEAS    : UDINT := 16#0005_0256; // 0005_0256 测量时长为零【故障级】/ Zero measure duration, fault level
    DL_LEAK_ERR_STATE   : UDINT := 16#0005_0257; // 0005_0257 非法状态兜底【故障级】/ Illegal state fallback, fault level
    DL_LEAK_INFO_LIMIT  : UDINT := 16#0005_0150; // 0005_0150 泄漏率上限为负，取绝对值【信息级】/ Negative leak limit, absolute taken, info level
    DL_LEAK_INFO_RISE   : UDINT := 16#0005_0151; // 0005_0151 测量窗压力回升（ΔP<0），按 0 处理【信息级】/ Pressure rise in window, floored, info level
    DL_LEAK_INFO_NOTC   : UDINT := 16#0005_0152; // 0005_0152 温度补偿已关闭，按原始压降判定【信息级】/ Temp compensation off, info level
    DL_LEAK_INFO_GROSS  : UDINT := 16#0005_0153; // 0005_0153 大漏快判触发（提前判 NG）【信息级】/ Gross-leak quick judge triggered, info level
END_VAR

// ============================================================================
// 段 1｜实例无条件周期刷新（R7/0.5：严禁置于 IF/CASE 分支内）
//      Unconditional per-cycle refresh of all instances (R7/0.5)
// ============================================================================
_fbTrigStart(CLK := bStart);            // 启动沿（Start edge）
_fbTrigReset(CLK := bReset);            // 复位沿（Reset edge）
_fbTonClampTo(IN := (_ePhase = E_DL_LeakPhase.eClampCheck), PT := tFillTimeout);  // 夹具确认超时（Clamp timeout）
_fbTonFillMin(IN := (_ePhase = E_DL_LeakPhase.eFill), PT := tFill);               // 最小充气保持（Min fill hold）
_fbTonFillTo(IN := (_ePhase = E_DL_LeakPhase.eFill), PT := tFillTimeout);         // 充气超时（Fill timeout）
_fbTonStab(IN := (_ePhase = E_DL_LeakPhase.eStabilize), PT := tStabilize);        // 稳压时长（Stabilize duration）
_fbTonMeas(IN := (_ePhase = E_DL_LeakPhase.eMeasure), PT := tMeasure);            // 测量时长（Measure duration）
_fbTonVentTo(IN := (_ePhase = E_DL_LeakPhase.eVent), PT := tVentTimeout);         // 排气超时（Vent timeout）

// 扫描周期秒值折算（R14：周期变更经相位切换自然断输入归零；此处每拍重算）
// Cycle seconds conversion (R14: phase switches naturally break timer input)
_fDtS := TIME_TO_REAL(tCycle) / DL_TIME_MS_SCALE;    // 毫秒 → 秒，本行换算单位为 s（Conversion unit: seconds）

// ============================================================================
// 段 2｜信息级预清零 + 输入防御 + 复位路径（R15）
//      Info preset + input defense + reset path (R15)
// ============================================================================
_uInfoCode := 0;                        // 信息级瞬时型每拍重算（Transient info recomputed each scan）
bDone := FALSE;                         // 判定单拍先清零（R25：置位-消费-复位同周期闭环）/ Done pulse preset FALSE (R25)

// 泄漏率上限负值取绝对值（Negative leak limit, absolute taken）
IF fLeakLimit < 0.0 THEN
    _fLeakLimEff := ABS(fLeakLimit);    // 取绝对值（Absolute value）
    _uInfoCode := DL_LEAK_INFO_LIMIT;   // 0005_0150 上限为负取绝对值【信息级】/ Negative limit, info level
ELSE
    _fLeakLimEff := fLeakLimit;         // 引脚原值（Pin value as-is）
END_IF

// REAL 输入非有限值/域防御（偏离留档①：tCycle 归并本码防御）
// REAL input non-finite/domain defense (deviation 1: tCycle folded into this code)
IF (NOT (fActPressure >= (-DL_LEAK_REAL_MAX) AND fActPressure <= DL_LEAK_REAL_MAX))
OR (NOT (fActTemp    >= (-DL_LEAK_REAL_MAX) AND fActTemp    <= DL_LEAK_REAL_MAX))
OR (NOT (fRefTemp    >= (-DL_LEAK_REAL_MAX) AND fRefTemp    <= DL_LEAK_REAL_MAX))
OR (NOT (fTestPressure >= (-DL_LEAK_REAL_MAX) AND fTestPressure <= DL_LEAK_REAL_MAX))
OR (NOT (fPressureTol  >= (-DL_LEAK_REAL_MAX) AND fPressureTol  <= DL_LEAK_REAL_MAX))
OR (NOT (fChamberVolume >= (-DL_LEAK_REAL_MAX) AND fChamberVolume <= DL_LEAK_REAL_MAX))
OR (NOT (fGrossLeakDrop >= (-DL_LEAK_REAL_MAX) AND fGrossLeakDrop <= DL_LEAK_REAL_MAX))
OR (NOT (fLeakLimit   >= (-DL_LEAK_REAL_MAX) AND fLeakLimit   <= DL_LEAK_REAL_MAX))
OR (NOT (tCycle >= T#1MS)) THEN
    _bFaultLatch := TRUE;               // 输入非有限值/周期非法锁存（Input defense latch）
    _uErrorIdInt := DL_LEAK_ERR_NAN;    // 0005_0254 输入非有限值【故障级】/ Non-finite input, fault level
    _ePhase := E_DL_LeakPhase.eFault;
ELSIF fChamberVolume <= 0.0 THEN
    _bFaultLatch := TRUE;               // 容积非法锁存（Volume defense latch）
    _uErrorIdInt := DL_LEAK_ERR_VOL;    // 0005_0255 腔容积非法【故障级】/ Invalid volume, fault level
    _ePhase := E_DL_LeakPhase.eFault;
ELSIF tMeasure = T#0MS THEN
    _bFaultLatch := TRUE;               // 测量时长为零锁存（Zero measure latch）
    _uErrorIdInt := DL_LEAK_ERR_MEAS;   // 0005_0256 测量时长为零【故障级】/ Zero measure duration, fault level
    _ePhase := E_DL_LeakPhase.eFault;
ELSE
    // 域钳位后的生效参数（Sanitized effective parameters）
    _fTestPressEff := LIMIT(DL_LEAK_PRESS_MIN, fTestPressure, DL_LEAK_PRESS_MAX); // 目标压力域钳位（Pressure clamped）
    _fTolEff       := LIMIT(DL_LEAK_TOL_MIN, fPressureTol, DL_LEAK_TOL_MAX);      // 容差域钳位（Tolerance clamped）
    _fVolEff       := fChamberVolume;   // 容积已过正数防御（Volume defended positive）
    _fGrossEff     := fGrossLeakDrop;   // 大漏阈（0=禁用快判）/ Gross threshold (0 = off)
END_IF

// 复位路径：仅此路径可清故障锁存与判定（R15）
IF _fbTrigReset.Q THEN
    _bFaultLatch := FALSE;              // 故障锁存解除（Fault latch released）
    _uErrorIdInt := 16#0000_0000;       // 故障码清零（Fault code cleared）
    _bAbortActive := FALSE;             // 中止锁存解除（Abort latch released）
    _bVerdictValid := FALSE;            // 判定失效（Verdict invalidated）
    _bPassLatched := FALSE;             // 判定锁存清零（Verdict latch cleared）
    IF _ePhase = E_DL_LeakPhase.eFault THEN
        _ePhase := E_DL_LeakPhase.eIdle; // 故障态回空闲（Fault phase back to idle）
    END_IF
END_IF

// ============================================================================
// 段 3｜中止电平全局拦截（优先级最高：任意执行相 → 安全排气）
//      Abort level global intercept (highest priority: safe vent from any active phase)
// ============================================================================
IF bAbort AND (NOT _bAbortActive)
AND (_ePhase <> E_DL_LeakPhase.eIdle) AND (_ePhase <> E_DL_LeakPhase.eFault)
AND (_ePhase <> E_DL_LeakPhase.ePass) AND (_ePhase <> E_DL_LeakPhase.eFail) THEN
    _bAbortActive := TRUE;              // 中止锁存（Abort latched）
    _bVerdictValid := FALSE;            // 判定作废不记 NG（Verdict voided, no NG recorded）
    _ePhase := E_DL_LeakPhase.eAbort;   // 进入安全排气（Enter safe vent）
END_IF

// ============================================================================
// 段 4｜核心相位状态机（ENUM + CASE，含 ELSE 非法状态兜底）
//      Core phase state machine (ENUM + CASE with ELSE fallback)
// ============================================================================
IF NOT bEnable THEN
    // 使能撤销：阀组安全侧（充气/隔离关、排气开）、判定清、相位回空闲
    // Disabled: valves to safe side, verdicts cleared, phase back to idle
    _ePhase := E_DL_LeakPhase.eIdle;
    _bVerdictValid := FALSE;
    _bPassLatched := FALSE;
    _bAbortActive := FALSE;
ELSE
    CASE _ePhase OF

        E_DL_LeakPhase.eIdle: // 空闲：等启动沿
            IF _fbTrigStart.Q AND (NOT _bFaultLatch) AND (NOT _bAbortActive) THEN
                _ePhase := E_DL_LeakPhase.eClampCheck;   // 受理启动（Start accepted）
            END_IF

        E_DL_LeakPhase.eClampCheck: // 夹具确认：等闭合信号
            IF bFixtureClosed THEN
                _ePhase := E_DL_LeakPhase.eFill;         // 夹具确认通过（Clamp confirmed）
            ELSIF _fbTonClampTo.Q THEN
                _bFaultLatch := TRUE;                    // 夹具未闭超时（Clamp timeout）
                _uErrorIdInt := DL_LEAK_ERR_CLAMP;       // 0005_0250 夹具闭合超时【故障级】/ Clamp timeout, fault level
                _ePhase := E_DL_LeakPhase.eFault;
            END_IF

        E_DL_LeakPhase.eFill: // 充气：最小保持到 + 压力达标双条件（偏离留档②）
            IF _fbTonFillMin.Q
            AND (fActPressure >= _fTestPressEff * (1.0 - DL_LEAK_FILL_TOL)) THEN
                _ePhase := E_DL_LeakPhase.eStabilize;    // 达标进稳压（Reached, stabilize）
            ELSIF _fbTonFillTo.Q THEN
                _bFaultLatch := TRUE;                    // 充气超时（Fill timeout）
                _uErrorIdInt := DL_LEAK_ERR_FILL;        // 0005_0251 充气超时未达压【故障级】/ Fill timeout, fault level
                _ePhase := E_DL_LeakPhase.eFault;
            END_IF

        E_DL_LeakPhase.eStabilize: // 稳压：隔离保温，结束时记录起点并判容差
            IF _fbTonStab.Q THEN
                _fP0 := fActPressure;                    // 测量起点压力（Pressure at start）
                _fT0 := fActTemp;                        // 测量起点温度（Temperature at start）
                _fMeasSec := 0.0;                        // 测量秒值累计清零（Measure seconds reset）
                IF ABS(_fP0 - _fTestPressEff) > _fTolEff THEN
                    _bFaultLatch := TRUE;                // 设备异常：稳压后压力超容差（Equipment fault: out of tolerance）
                    _uErrorIdInt := DL_LEAK_ERR_STAB;    // 0005_0252 稳压超容差（不判工件 NG）【故障级】/ Stabilize out of tolerance, equipment fault
                    _ePhase := E_DL_LeakPhase.eFault;
                ELSE
                    _ePhase := E_DL_LeakPhase.eMeasure;  // 进入隔离测量（Enter measure）
                END_IF
            END_IF

        E_DL_LeakPhase.eMeasure: // 测量：实时压差跟踪 + 大漏快判 + 计时结算
            _fMeasSec := _fMeasSec + _fDtS;              // 测量秒值累计（Measure seconds accumulate）
            _fDeltaPInt := _fP0 - fActPressure;          // 实时压差（Live delta-P）
            IF _fDeltaPInt < 0.0 THEN
                _fDeltaPInt := 0.0;                      // 压力回升按 0 处理（Rise floored to zero）
                _uInfoCode := DL_LEAK_INFO_RISE;         // 0005_0151 压力回升【信息级】/ Pressure rise, info level
            END_IF
            IF (_fGrossEff > 0.0) AND (_fDeltaPInt >= _fGrossEff) THEN
                _uInfoCode := DL_LEAK_INFO_GROSS;        // 0005_0153 大漏快判触发【信息级】/ Gross-leak quick judge, info level
                fDeltaP := _fDeltaPInt;                 // 压差锁存（Delta-P latched）
                fLeakRate := 0.0;                        // 快判路径无有效泄漏率（No rate on gross path）
                _bPassLatched := FALSE;                  // 不合格锁存（Fail latched）
                _bVerdictValid := TRUE;
                nPartCount := nPartCount + UINT#1;       // 计件（Part counted）
                nRejectCount := nRejectCount + UINT#1;   // 计不良（Reject counted）
                bDone := TRUE;                           // 判定单拍（R25 本拍闭环）/ Done pulse (R25)
                _ePhase := E_DL_LeakPhase.eVent;
            ELSIF _fbTonMeas.Q THEN
                // 测量窗到期结算（Measure window settled）
                fDeltaP := _fDeltaPInt;                 // 压差锁存（Delta-P latched）
                IF _fMeasSec > DL_LEAK_EPS THEN
                    _fLeakRateInt := _fDeltaPInt * _fVolEff / _fMeasSec * DL_LEAK_UNIT_FACTOR;
                    // 量纲链：kPa·mL/s × 60 → mL/min（偏离留档②前的设计要点④完整推导）
                    // Unit chain: kPa*mL/s times 60 = mL/min (full derivation in key notes 4)
                ELSE
                    _fLeakRateInt := 0.0;                // 秒值防御（除零保护，理论上不可达）/ Divide guard (unreachable by design)
                END_IF
                IF bTempCompEnable THEN
                    _fDenK := DL_LEAK_KELVIN + _fT0;     // 补偿分母（Compensation denominator）
                    IF _fDenK > DL_LEAK_EPS THEN
                        _fLeakRateInt := _fLeakRateInt * (DL_LEAK_KELVIN + fRefTemp) / _fDenK;
                        // 一阶理想气体近似（设计要点④声明适用域）/ First-order ideal-gas approximation
                    END_IF
                ELSE
                    _uInfoCode := DL_LEAK_INFO_NOTC;     // 0005_0152 温度补偿关闭【信息级】/ Temp compensation off, info level
                END_IF
                fLeakRate := _fLeakRateInt;              // 泄漏率锁存（Rate latched）
                _bPassLatched := _fLeakRateInt <= _fLeakLimEff;  // 判定：≤ 上限为合格（Verdict by limit）
                _bVerdictValid := TRUE;
                nPartCount := nPartCount + UINT#1;       // 计件（Part counted）
                IF NOT _bPassLatched THEN
                    nRejectCount := nRejectCount + UINT#1;   // 计不良（Reject counted）
                END_IF
                bDone := TRUE;                           // 判定单拍（R25 本拍闭环）/ Done pulse (R25)
                _ePhase := E_DL_LeakPhase.eVent;
            END_IF

        E_DL_LeakPhase.eVent: // 排气：泄压到安全位后分流（中止→空闲 / 判定→保持态）
            IF fActPressure < DL_LEAK_VENT_DONE THEN
                IF _bAbortActive THEN
                    _bAbortActive := FALSE;              // 中止路径排气完成回空闲（Abort vent done back to idle）
                    _ePhase := E_DL_LeakPhase.eIdle;
                ELSIF _bVerdictValid THEN
                    // 正常判定路径排气完成后进保持态（Verdict hold phase after vent done）
                    IF _bPassLatched THEN
                        _ePhase := E_DL_LeakPhase.ePass; // 合格保持（Pass hold）
                    ELSE
                        _ePhase := E_DL_LeakPhase.eFail; // 不合格保持（Fail hold）
                    END_IF
                ELSE
                    _ePhase := E_DL_LeakPhase.eIdle;     // 无判定兜底回空闲（No verdict, back to idle）
                END_IF
            ELSIF _fbTonVentTo.Q THEN
                _bFaultLatch := TRUE;                    // 排气超时（Vent timeout）
                _uErrorIdInt := DL_LEAK_ERR_VENT;        // 0005_0253 排气超时【故障级】/ Vent timeout, fault level
                _ePhase := E_DL_LeakPhase.eFault;
            END_IF

        E_DL_LeakPhase.ePass: // 合格保持：等复位或新周期
            IF _fbTrigStart.Q AND (NOT _bFaultLatch) AND (NOT bAbort) THEN
                _ePhase := E_DL_LeakPhase.eClampCheck;   // 新周期受理（New cycle accepted）
                _bVerdictValid := FALSE;
                bPass := FALSE;
            END_IF

        E_DL_LeakPhase.eFail: // 不合格保持：等复位或新周期
            IF _fbTrigStart.Q AND (NOT _bFaultLatch) AND (NOT bAbort) THEN
                _ePhase := E_DL_LeakPhase.eClampCheck;   // 新周期受理（New cycle accepted）
                _bVerdictValid := FALSE;
                bFail := FALSE;
            END_IF

        E_DL_LeakPhase.eAbort: // 中止排气：泄压到安全位后保持等待复位
            IF fActPressure < DL_LEAK_VENT_DONE THEN
                _bAbortActive := FALSE;                  // 安全位达成，中止释放（Safe level reached, abort released）
            END_IF

        E_DL_LeakPhase.eFault: // 设备故障锁存：等复位（复位路径在段 2）
            // 等复位（Awaiting reset）

        ELSE // 非法状态兜底（本块专用码位）
            _bFaultLatch := TRUE;
            _uErrorIdInt := DL_LEAK_ERR_STATE;           // 0005_0257 非法状态兜底【故障级】/ Illegal state fallback, fault level
            _ePhase := E_DL_LeakPhase.eFault;
    END_CASE
END_IF

// 复位路径补充：保持态复位回空闲（Hold phases reset back to idle）
IF _fbTrigReset.Q AND ((_ePhase = E_DL_LeakPhase.ePass) OR (_ePhase = E_DL_LeakPhase.eFail)) THEN
    _ePhase := E_DL_LeakPhase.eIdle;     // 保持态复位（Hold released）
END_IF

// ============================================================================
// 段 5｜输出派生（阀组安全侧 + 判定互斥先清后置）
//      Output derivation (valve safe side + verdict mutual exclusion)
// ============================================================================
// 阀组默认安全侧：全关（Valves preset closed）
bCmdFillValve := FALSE;                  // 充气阀预清（Fill preset）
bCmdIsolateValve := FALSE;               // 隔离阀预清（Isolate preset）
bCmdVentValve := FALSE;                  // 排气阀预清（Vent preset）

IF bEnable AND (NOT _bFaultLatch) THEN
    bCmdFillValve := (_ePhase = E_DL_LeakPhase.eFill);          // 充气阀：仅充气相（Fill in fill phase）
    bCmdIsolateValve := (_ePhase = E_DL_LeakPhase.eStabilize)
                     OR (_ePhase = E_DL_LeakPhase.eMeasure);    // 隔离阀：稳压与测量相（测量前必须隔离气源）/ Isolate in stabilize+measure
    bCmdVentValve := (_ePhase = E_DL_LeakPhase.eVent)
                  OR (_ePhase = E_DL_LeakPhase.eAbort)
                  OR _bAbortActive;                             // 排气阀：排气/中止相与中止锁存期（Vent in vent/abort）
ELSE
    bCmdVentValve := TRUE;               // 使能撤销/故障：安全排气（Safe vent on disable or fault）
END_IF

// 判定互斥先清后置（出口断言：bPass 与 bFail 恒互斥）
// Verdict mutual exclusion: preset clear then set (exit assertion)
bPass := FALSE;                          // 合格预清（Pass preset）
bFail := FALSE;                          // 不合格预清（Fail preset）
IF _bVerdictValid THEN
    bPass := _bPassLatched;              // 合格出口（Pass outlet）
    bFail := NOT _bPassLatched;          // 不合格出口（Fail outlet）
END_IF

bBusy := (_ePhase = E_DL_LeakPhase.eClampCheck)
      OR (_ePhase = E_DL_LeakPhase.eFill)
      OR (_ePhase = E_DL_LeakPhase.eStabilize)
      OR (_ePhase = E_DL_LeakPhase.eMeasure)
      OR (_ePhase = E_DL_LeakPhase.eVent);               // 周期执行中派生（Busy derived）

ePhase := _ePhase;                       // 相位镜像（Phase mirror）

// ============================================================================
// 段 6｜bError/uErrorId 出口（R21：bError 显式排除信息级码）
//      Outlets: bError excludes info codes (R21)
// ============================================================================
bError := _bFaultLatch;                  // 故障级派生式（Fault-level derived form）
IF _bFaultLatch THEN
    uErrorId := _uErrorIdInt;            // 故障级码优先透出（Fault-level priority）
ELSE
    uErrorId := _uInfoCode;              // 无故障时透出本拍信息级码（Transient info code）
END_IF
END_FUNCTION_BLOCK

(* ---- FB_DL_MixRecipeControl.st ---- *)
(*==============================================================================
 * 组件名称 (Component)  : FB_DL_MixRecipeControl
 * 所属子库 (Sublibrary) : DL_Process
 * 当前版本 (Version)    : 1.0.1
 * 兼容性 (Platform)   : CODESYS 3.5 / TwinCAT 3 / 汇川 InoProShop / Machine Expert
 *                         仅依赖 Standard.library（TON / R_TRIG）+ 既有接口
 *                         I_DL_VfdDrive（DL_Device R6 契约件，仅引用零修改）
 * 分类     (Category)   : 工艺段功能块（Function Block · ISA-88 单相语义混合搅拌）
 * 功能简述 (Function)   : 混合/搅拌工艺相控制（ISA-88 单相语义 clean-room）：
 *                         投料就绪 → 搅拌（定速/正反交替）→ 终点判据（时间
 *                         到/扭矩上升达标）→ 出料许可 → 停转；转速反馈监视、
 *                         扭矩超限保护、出料超时诊断。驱动控制全部经 I_DL_Vfd
 *                         Drive 接口引用（引脚注入），本块零硬件依赖。
 * 接口消费 (Consumes)   : I_DL_VfdDrive（既有契约，仅引用零修改）：每拍至多
 *                         一次方法调用（公约 0.13），由内部单发指令调度器串行
 *                         化——CmdStop > CmdRun > SetFrequency 优先级链；接
 *                         口无 bReady 属性，前置就绪按 NOT iDrive.bFault 判
 *                         定（R11 留档见偏离留档①）；SetFrequency 引脚值域
 *                         为 Hz，本块传入转速数值，rpm↔Hz 标定由调用方实现
 *                         块承担（既有契约语义，头注释声明）。
 * 首扫说明 (Init note)  : 顺序型组件但全部状态由指令沿/电平驱动，免首扫
 *                         （R23/公约 0.1），无 bInit。
 * 公约遵循 (Convention) : 0.2/R21 bError 仅故障级码置位；0.4 双语同行注释；
 *                         0.5/R7 实例主体最前部无条件刷新；0.7/R15 故障锁存
 *                         仅复位路径清码；0.10 定时基准由引脚给（tCycle 增补
 *                         引脚，泳道 A 同款公共约定，非逐组件条款）；0.13 接
 *                         口调用配额每拍至多一次（调度器结构保证）；0.14 非
 *                         有限值防御；0.15 转速统一 rpm、扭矩统一 % 额定；
 *                         0.16 无魔法数；0.17 终结符成对 ✓；0.19 码位同行
 *                         【级别】注释；0.20 验收向量入头注释；R25 bDone 单
 *                         拍三律。
 * 红线自检 (Redline)    : R1 零全局变量表/外部变量引用 ✓｜R2 零物理 IO 地址 ✓
 *                         R3 纯 IEC 61131-3 ✓｜R4 非有限值/除零/浮点容差 ✓
 *                         R5 全变量中英双语同行注释 ✓｜R6 ENUM+CASE+ELSE ✓
 *                         R7 五实例（R_TRIG×2/TON×3）主体最前部无条件刷新 ✓
 *                         R8 全常量化 ✓｜R25 单拍标志生命周期三律 ✓
 * 设计要点 (Key notes)  : ① 接口单发调度器：状态机只登记指令请求标志，唯一
 *                           的方法调用点在段 6 调度器（Stop > Run > SetFreq
 *                           优先级链），结构上保证每拍至多一次方法调用（公约
 *                           0.13）；SetFrequency 仅在设定变化超容差时下发；
 *                         ② 交替换向三步序（禁止直接反接，防机械冲击）：
 *                           CmdStop → 等 fActSpeed < DL_MIX_STOP_EPS →
 *                           CmdRun(新方向) → 下一拍补发 SetFrequency；
 *                         ③ 转速确认窗：进入搅拌相后 tSpeedCheck 内须达 90%
 *                           设定，否则 0261（皮带断/驱动未使能类故障）；混合
 *                           计时仅在确认通过后累计（暂停期冻结）；
 *                         ④ 扭矩保护：fActTorque ≥ fTorqueLimit 立即停 + 故
 *                           障 0263（疑似卡桨/物料过稠，防烧电机）；
 *                         ⑤ 方向互斥出口断言：bDirForward 与 bDirReverse 由
 *                           同一方向寄存器派生，结构上恒互斥（切换过渡期双
 *                           FALSE）；
 *                         ⑥ fProgress 量纲推导：已混合秒值/目标秒值 [-]，双
 *                           方经 TIME 毫秒口径转 REAL 后相除（除前判零），钳
 *                           位 [0,1]。
 * 偏离留档 (Deviation)  : 依 R11 头注释留档，共 2 条：
 *                         ① 前置就绪判据：规格预留「若接口无 bReady 属性改
 *                           用 NOT iDrive.bFault」——既有 I_DL_VfdDrive 契
 *                           约无 bReady，本块按 NOT iDrive.bFault 实现，规格
 *                           预案内非语义偏离；
 *                         ② tCycle 增补引脚：混合计时累计与进度折算需要时
 *                           间基准，依公约 0.10 增补（泳道 A 先例，公共约定
 *                           强制项，非逐组件条款）。
 * 开源溯源 (Origin)     : 来源标签 isa-88-phase / mixing-process（RAW_NOTES_R8
 *                         S-9 LBP 实测 + S-10 相语义：ISA-88 相（Phase）公开
 *                         语义——前确认/执行/终点判据/完成的相结构与「批次数
 *                         据不进控制逻辑」的分层思想，公开技术资料，仅借鉴相
 *                         分类与参数域；状态机、交替换向三步序、码位、引脚契
 *                         约 100% 本库独立设计，clean-room 未复制源码。许可
 *                         证说明：ISA-88 为公开标准语义，本文件为本库原创实
 *                         现，随本库许可证发布）。
 * 验收向量 (Acceptance) :
 *   V1 正常混合 tMixTime → bOk + bDone 单拍 + fProgress≈1.0；
 *   V2 交替模式（30 s 换向）：方向互斥、先停后启无直接反接；
 *   V3 扭矩超限 → 立即停 + 故障 0263；
 *   V4 转速确认窗内未建立 → 0261；
 *   V5 bEndByTorque 且扭矩提前达标 → 信息码 0163 提前完成；
 *   V6 超最长混合时间 → eNg + 信息码 0162；
 *   V7 出料超时 → 0262；
 *   V8 bAbort 中途 → 停转且不出料、无 OK/NG。
 * 修订历史 (Revision)   :
 *   2026-11-15  v1.0.0  首版入库（Round 08 · DL_Process 混合工艺相件）
 *   2026-11-15  v1.0.1  R8 总监终审修复四项：① eMixing 判 NG 分支写入未声明
 *                       内部变量 _bNg（编译期未定义符号）改为出口 bNg；② 判
 *                       定保持语义补齐——eDone 相每拍置 bOk、eNg 相每拍置 bNg
 *                       （原仅转换拍脉冲，违反规格「eDone/eNg 保持」）；③ 最
 *                       长混合时间判据与目标时间判据的 ELSIF 先后倒置导致
 *                       eNg 终态不可达（tElapsed ≥ tMixMax 必先被 tElapsed ≥
 *                       tMixEff 捕获），改为「扭矩终点 → 时间模式目标终点 →
 *                       最长超时」序，恢复 V6 可达性且时间模式无回归；④ 终端
 *                       态分支内孤立空语句 `;`（非 IEC 61131-3 文法）改为纯注
 *                       释占位分支。
 *============================================================================*)

(*-----------------------------------------------------------------------------
 * 枚举: E_DL_MixPhase（归属 FB_DL_MixRecipeControl，与其同文件发布，公约 0.18）
 *----------------------------------------------------------------------------*)
TYPE E_DL_MixPhase :
(
    eIdle      := 0,   // 空闲：等启动 / Idle, awaiting start
    ePreCheck  := 10,  // 前置确认：料已投、出料阀关、驱动就绪 / Precheck, material, outlet and drive ready
    eMixing    := 20,  // 搅拌中（含交替子计时）/ Mixing with alternate sub-timing
    eVerify    := 30,  // 终点确认：稳速确认与结果锁存 / Verify, speed stability and result latch
    eDischarge := 40,  // 出料中：等出料完成信号 / Discharging, awaiting discharge done
    eSpinDown  := 50,  // 停转：减速到零 / Spin down to standstill
    eDone      := 60,  // 完成（OK），等复位 / Done, awaiting reset
    eNg        := 70,  // 不合格（终点未达但超最长混合时间），等复位 / NG on max-time expiry, awaiting reset
    eAbort     := 80,  // 中止：立即停转，禁止出料 / Aborted, stopped and discharge forbidden
    eFault     := 99   // 故障锁存 / Fault latched
) UINT;
END_TYPE

FUNCTION_BLOCK FB_DL_MixRecipeControl
VAR_INPUT
    bEnable             : BOOL;             // 使能（Enable），FALSE=停转清输出 / Enable, FALSE stops drive and clears outputs
    bStart              : BOOL;             // 启动混合相（Start），上升沿受理（空闲/完成/不合格态）/ Start edge accepted at idle/done/ng
    bAbort              : BOOL;             // 中止（Abort），电平最高优先：停转、禁止出料 / Abort level, highest priority
    bReset              : BOOL;             // 复位（Reset），上升沿受理 / Rising edge resets fault and verdicts
    bMaterialReady      : BOOL;             // 投料就绪（Material ready），前置确认项 / Material loaded interlock
    bOutletClosed       : BOOL;             // 出料阀关闭确认（Outlet closed），前置确认项 / Outlet valve closed interlock
    bDischargeDone      : BOOL;             // 出料完成（Discharge done），出料相退出条件 / Discharge completion feedback
    fSpeedSetpoint      : REAL := 300.0;    // 搅拌转速设定（Speed setpoint）[rpm]，域 1..3000，越界钳位 / Speed setpoint [rpm]
    fActSpeed           : REAL;             // 实际转速（Actual speed）[rpm]，由变频器/适配层注入 / Actual speed [rpm] injected
    fActTorque          : REAL;             // 实际扭矩（Actual torque）[% 额定] / Actual torque [% of rated]
    fTorqueLimit        : REAL := 85.0;     // 扭矩保护上限（Torque limit）[%]，超限即停 + 故障 / Torque protection limit [%]
    bEndByTorque        : BOOL;             // 以扭矩上升为终点判据（End by torque），TRUE=扭矩达标即完成 / Torque-rise end criterion enable
    fTorqueRiseTarget   : REAL := 60.0;     // 终点扭矩判据（End torque target）[%]，仅 bEndByTorque 有效 / Torque end target [%]
    tMixTime            : TIME := T#5M;     // 目标混合时间（Mix time）/ Target mix duration
    tMixTimeMax         : TIME := T#15M;    // 最长混合时间（Max mix time），超时判 NG / Maximum mix duration, expiry = NG
    bAlternate          : BOOL;             // 正反交替（Alternate direction），TRUE=每 tAlternateTime 换向 / Alternate direction enable
    tAlternateTime      : TIME := T#30S;    // 交替周期（Alternate period），仅 bAlternate 有效 / Alternate period
    tSpeedCheck         : TIME := T#5S;     // 转速到位确认窗（Speed check window），窗内须达 90% 设定 / Speed establish window
    tDischargeTimeout   : TIME := T#60S;    // 出料超时（Discharge timeout）/ Discharge timeout
    tCycle              : TIME := T#10MS;   // 任务扫描周期（Task cycle time）[ms]，由调用方按实际任务给，计时累计基准（公约 0.10）/ Task cycle time, timing base
END_VAR
VAR_OUTPUT
    fSpeedCmd           : REAL;             // 转速指令（Speed command）[rpm]，0=停 / Speed command [rpm], zero = stop
    bDirForward         : BOOL;             // 正转指令（Forward），与反转互斥 / Forward direction, exclusive with reverse
    bDirReverse         : BOOL;             // 反转指令（Reverse）/ Reverse direction
    ePhase              : E_DL_MixPhase := E_DL_MixPhase.eIdle; // 当前相位（Current phase）/ Current phase
    bBusy               : BOOL;             // 执行中（Busy），前置确认至停转态为 TRUE / TRUE from precheck to spin-down
    bDone               : BOOL;             // 完成单拍脉冲（Done pulse，OK 或 NG 进入时各一次），单拍生命周期三律 / One-scan verdict pulse
    bOk                 : BOOL;             // 混合合格（OK），完成保持态为 TRUE / OK verdict held
    bNg                 : BOOL;             // 混合不合格（NG），不合格保持态为 TRUE / NG verdict held
    fProgress           : REAL;             // 进度（Progress）[-]，0.0..1.0 = 已混合时间/目标时间（钳位）/ Mix progress dimensionless clamped
    tElapsed            : TIME := T#0S;     // 已混合时长（Elapsed mix time），仅确认通过后累计 / Elapsed mix time, accumulates after confirm
    bError              : BOOL;             // 故障锁存（Error），仅故障级码 / Latched error, fault codes only
    uErrorId            : UDINT;            // 故障码（Error code），16#0005_xxxx 段，0=无故障 / Error code, fault-level priority
END_VAR
VAR_IN_OUT
    iDrive              : I_DL_VfdDrive;    // 搅拌驱动接口引用（Mixer drive，既有契约 I_DL_VfdDrive），由上层注入实例 / Mixer drive interface reference injected by caller
END_VAR
VAR
    _ePhase             : E_DL_MixPhase := E_DL_MixPhase.eIdle;   // 内部相位（Internal phase）/ Internal phase
    _bFaultLatch        : BOOL;             // 故障锁存标志（Fault latch flag），仅复位路径清除 / Fault latch, cleared only via reset path
    _uErrorIdInt        : UDINT;            // 内部故障级码寄存（Internal fault-level register）/ Internal fault-level register
    _uInfoCode          : UDINT;            // 本拍信息级码（Info code this cycle），瞬时型每拍重算 / Transient info code
    _bCmdStopReq        : BOOL;             // 停止指令请求（Stop request flag），调度器消费 / Stop request consumed by dispatcher
    _bCmdRunReq         : BOOL;             // 运行指令请求（Run request flag），调度器消费 / Run request consumed by dispatcher
    _bCmdFreqReq        : BOOL;             // 频率设定请求（Frequency request flag），调度器消费 / Frequency request consumed by dispatcher
    _bRunFwd            : BOOL;             // 待发方向（Pending direction），TRUE=正转 / Pending direction, TRUE = forward
    _bRunIssued         : BOOL;             // 运行指令已受理锁存（Run accepted latch）/ Run accepted latch
    _bDirFwd            : BOOL := TRUE;     // 当前方向寄存（Current direction register），TRUE=正转 / Current direction, TRUE = forward
    _bConfirmed         : BOOL;             // 转速确认通过（Speed confirmed）/ Speed establish confirmed
    _bRevPending        : BOOL;             // 换向请求（Reversal pending）/ Reversal pending
    _bRevInStop         : BOOL;             // 换向停转步（Reversal stop step），等待转速落零 / Reversal stop step, waiting speed near zero
    _tElapsedInt        : TIME := T#0S;     // 内部混合计时（Internal mix elapsed），确认后每拍加 tCycle / Internal elapsed, accumulates after confirm
    _fSetEff            : REAL;             // 生效转速设定（Effective setpoint）[rpm]，钳位后值 / Sanitized setpoint [rpm]
    _fTorqueLimEff      : REAL;             // 生效扭矩上限（Effective torque limit）[%] / Sanitized torque limit [%]
    _fTorqueTgtEff      : REAL;             // 生效终点扭矩（Effective end torque target）[%] / Sanitized end torque target [%]
    _tMixEff            : TIME;             // 生效目标混合时间（Effective mix time）/ Sanitized mix duration
    _tMixMaxEff         : TIME;             // 生效最长混合时间（Effective max mix time）/ Sanitized max mix duration
    _tAltEff            : TIME;             // 生效交替周期（Effective alternate period）/ Sanitized alternate period
    _tAltLast           : TIME := T#30S;    // 上拍生效交替周期（Last alternate period），PT 变更检测基准 / Last alternate period for PT-change detection
    _bAltBreak          : BOOL := TRUE;     // 交替计时输入使能（Alternate input enable），PT 变更拍断一拍 / Alternate input enable, broken on PT change
    _fFreqReq           : REAL;             // 待发频率值（Pending frequency value），调度器消费 / Pending frequency value
    _fFreqLast          : REAL;             // 末次下发频率（Last sent frequency），变化超容差才重发 / Last sent frequency, resend on change
    _fSpeedCmdInt       : REAL;             // 内部转速指令（Internal speed command）[rpm] / Internal speed command [rpm]
    _bFiniteSpd         : BOOL;             // 转速信号有限（Speed finite verdict）/ Speed signal finite verdict
    _bFiniteTrq         : BOOL;             // 扭矩信号有限（Torque finite verdict）/ Torque signal finite verdict
    _fbTrigStart        : R_TRIG;           // 启动沿（Start edge detector）/ Start edge detector
    _fbTrigReset        : R_TRIG;           // 复位沿（Reset edge detector）/ Reset edge detector
    _fbTonPreChk        : TON;              // 前置确认窗（Precheck window）/ Precheck window timer
    _fbTonSpdChk        : TON;              // 转速确认窗（Speed establish window）/ Speed establish window timer
    _fbTonAlt           : TON;              // 交替周期（Alternate period）/ Alternate period timer
    _fbTonDischTo       : TON;              // 出料超时（Discharge timeout）/ Discharge timeout timer
END_VAR
VAR CONSTANT
    DL_MIX_REAL_MAX     : REAL := 3.4E38;   // 单精度有限值判据幅值（Finite magnitude bound）/ Finite magnitude bound for REAL inputs
    DL_MIX_EPS          : REAL := 1.0E-6;   // 浮点防零/防重发容差（Float divide-guard epsilon）/ Float epsilon
    DL_MIX_STOP_EPS     : REAL := 1.0;      // 停转判定阈（Standstill threshold）[rpm]，低于此值视为已停 / Standstill speed threshold [rpm]
    DL_MIX_FREQ_EPS     : REAL := 0.5;      // 频率重发容差（Frequency resend epsilon）[rpm]，变化超此值才下发 / Resend threshold for setpoint change
    DL_MIX_SPD_OK_FRAC  : REAL := 0.9;      // 确认转速比例（Confirm speed fraction）[-]，达设定 90% 视为建立 / Confirm at 90% of setpoint
    DL_MIX_VERIFY_FRAC  : REAL := 0.05;     // 终点稳速容差比例（Verify tolerance fraction）[-]，±5% 设定 / Verify within 5% of setpoint
    DL_MIX_DISCHARGE_SPD: REAL := 50.0;     // 出料助排慢速（Discharge assist speed）[rpm] / Slow discharge assist speed [rpm]
    DL_MIX_SPD_MIN      : REAL := 1.0;      // 转速设定域下限（Setpoint lower clamp）[rpm] / Setpoint lower clamp [rpm]
    DL_MIX_SPD_MAX      : REAL := 3000.0;   // 转速设定域上限（Setpoint upper clamp）[rpm] / Setpoint upper clamp [rpm]
    DL_MIX_ALT_FACTOR   : DINT := 2;        // 交替周期提升倍数（Alternate raise factor）[-]，提升到确认窗的此倍数 / Alternate raise factor over check window
    DL_MIX_ERR_PRECHK   : UDINT := 16#0005_0260; // 0005_0260 前置条件不成立（料/阀/驱动）【故障级】/ Precheck timeout, fault level
    DL_MIX_ERR_SPEED    : UDINT := 16#0005_0261; // 0005_0261 转速未在确认窗内建立【故障级】/ Speed not established, fault level
    DL_MIX_ERR_DISCH    : UDINT := 16#0005_0262; // 0005_0262 出料超时【故障级】/ Discharge timeout, fault level
    DL_MIX_ERR_TORQUE   : UDINT := 16#0005_0263; // 0005_0263 扭矩超保护上限（疑似卡桨）【故障级】/ Torque over protection limit, fault level
    DL_MIX_ERR_NAN      : UDINT := 16#0005_0264; // 0005_0264 转速/扭矩信号非有限值【故障级】/ Non-finite speed or torque, fault level
    DL_MIX_ERR_STATE    : UDINT := 16#0005_0265; // 0005_0265 非法状态兜底【故障级】/ Illegal state fallback, fault level
    DL_MIX_INFO_CLAMP   : UDINT := 16#0005_0160; // 0005_0160 转速设定越界钳位【信息级】/ Setpoint clamped, info level
    DL_MIX_INFO_SWAP    : UDINT := 16#0005_0161; // 0005_0161 混合时间与最长混合时间对调自修复【信息级】/ Mix times swapped, info level
    DL_MIX_INFO_MAXT    : UDINT := 16#0005_0162; // 0005_0162 最长混合时间到，判 NG【信息级】/ Max mix time reached, NG, info level
    DL_MIX_INFO_TORQEND : UDINT := 16#0005_0163; // 0005_0163 以扭矩上升为终点判据触发【信息级】/ Torque-rise end criterion, info level
    DL_MIX_INFO_ALTRAISE: UDINT := 16#0005_0164; // 0005_0164 交替周期被提升至两倍确认窗【信息级】/ Alternate period raised, info level
END_VAR

// ============================================================================
// 段 1｜实例无条件周期刷新（R7/0.5：严禁置于 IF/CASE 分支内）
//      Unconditional per-cycle refresh of all instances (R7/0.5)
// ============================================================================
_fbTrigStart(CLK := bStart);            // 启动沿（Start edge）
_fbTrigReset(CLK := bReset);            // 复位沿（Reset edge）
_fbTonPreChk(IN := (_ePhase = E_DL_MixPhase.ePreCheck), PT := tSpeedCheck);   // 前置确认窗（Precheck window）
_fbTonSpdChk(IN := (_ePhase = E_DL_MixPhase.eMixing) AND (NOT _bConfirmed), PT := tSpeedCheck); // 转速确认窗（Speed window）
_fbTonAlt(IN := (_ePhase = E_DL_MixPhase.eMixing) AND _bConfirmed AND bAlternate
          AND (NOT _bRevPending) AND (NOT _bRevInStop) AND _bAltBreak, PT := _tAltEff);  // 交替周期（Alternate period）
_fbTonDischTo(IN := (_ePhase = E_DL_MixPhase.eDischarge), PT := tDischargeTimeout); // 出料超时（Discharge timeout）

// 交替周期 PT 变更断输入一拍（R14：防改时间常数后计时不清零的幽灵故障）
// Alternate-period PT-change one-scan input break (R14)
IF _tAltEff <> _tAltLast THEN
    _bAltBreak := FALSE;                // 交替计时输入断一拍（Alternate input broken one scan）
    _tAltLast := _tAltEff;              // 登记新交替周期（Register new alternate period）
ELSE
    _bAltBreak := TRUE;                 // 恢复交替计时输入（Alternate input restored）
END_IF

// ============================================================================
// 段 2｜信息级预清零 + 出口默认赋值（0.9：任何早退路径输出确定）+ 参数防御
//      Info preset + output defaults + parameter defense
// ============================================================================
_uInfoCode := 0;                        // 信息级瞬时型每拍重算（Transient info recomputed each scan）
bDone := FALSE;                         // 完成单拍先清零（R25：置位-消费-复位同周期闭环）/ Done pulse preset FALSE (R25)
fSpeedCmd := 0.0;                       // 转速指令默认停（Speed command default stop）
bDirForward := FALSE;                   // 方向默认双 FALSE（Directions default FALSE）
bDirReverse := FALSE;
bOk := FALSE;                           // 判定默认清（Verdicts preset）
bNg := FALSE;
fProgress := 0.0;                       // 进度默认零（Progress default zero）

// 信号非有限值防御（转速/扭矩，任何执行态均监视）
// Non-finite defense on speed/torque signals
_bFiniteSpd := (fActSpeed  >= (-DL_MIX_REAL_MAX)) AND (fActSpeed  <= DL_MIX_REAL_MAX);
_bFiniteTrq := (fActTorque >= (-DL_MIX_REAL_MAX)) AND (fActTorque <= DL_MIX_REAL_MAX);
IF bEnable AND ((NOT _bFiniteSpd) OR (NOT _bFiniteTrq)) THEN
    _bFaultLatch := TRUE;               // 信号非有限值锁存（Signal defense latch）
    _uErrorIdInt := DL_MIX_ERR_NAN;     // 0005_0264 转速/扭矩非有限值【故障级】/ Non-finite signal, fault level
    _ePhase := E_DL_MixPhase.eFault;
END_IF

// 转速设定钳位（Setpoint clamp，域 1..3000）
IF (fSpeedSetpoint < DL_MIX_SPD_MIN) OR (fSpeedSetpoint > DL_MIX_SPD_MAX) THEN
    _fSetEff := LIMIT(DL_MIX_SPD_MIN, fSpeedSetpoint, DL_MIX_SPD_MAX);   // 域钳位（Domain clamp）
    _uInfoCode := DL_MIX_INFO_CLAMP;    // 0005_0160 设定越界钳位【信息级】/ Setpoint clamped, info level
ELSE
    _fSetEff := fSpeedSetpoint;         // 引脚原值（Pin value as-is）
END_IF

// 混合时间与最长混合时间对调自修复（对调后目标 ≤ 上限）
// Mix times swap self-repair (target ≤ max after swap)
IF tMixTime > tMixTimeMax THEN
    _tMixEff := tMixTimeMax;            // 对调：目标取原上限（Swap: target = old max）
    _tMixMaxEff := tMixTime;            // 对调：上限取原目标（Swap: max = old target）
    _uInfoCode := DL_MIX_INFO_SWAP;     // 0005_0161 时间对调自修复【信息级】/ Times swapped, info level
ELSE
    _tMixEff := tMixTime;               // 引脚原值（Pin values as-is）
    _tMixMaxEff := tMixTimeMax;
END_IF

// 交替周期自动提升：小于两倍确认窗时提升到两倍（防换向太频转速永远建不起来）
// Alternate period auto-raise below twice check window (prevents never-established speed)
IF tAlternateTime < tSpeedCheck * DL_MIX_ALT_FACTOR THEN
    _tAltEff := tSpeedCheck * DL_MIX_ALT_FACTOR;    // 提升到两倍确认窗（Raised to twice window）
    _uInfoCode := DL_MIX_INFO_ALTRAISE;             // 0005_0164 交替周期被提升【信息级】/ Alternate raised, info level
ELSE
    _tAltEff := tAlternateTime;         // 引脚原值（Pin value as-is）
END_IF

// 扭矩限/终点扭矩防御（非有限值/非正回默认语义域钳位）
// Torque limit/target defense
_fTorqueLimEff := LIMIT(DL_MIX_EPS, fTorqueLimit, DL_MIX_REAL_MAX);        // 上限域钳位（Limit clamped）
_fTorqueTgtEff := LIMIT(DL_MIX_EPS, fTorqueRiseTarget, _fTorqueLimEff);    // 终点目标不超过保护上限（Target ≤ limit）

// 复位路径：仅此路径可清故障锁存与判定（R15）
IF _fbTrigReset.Q THEN
    _bFaultLatch := FALSE;              // 故障锁存解除（Fault latch released）
    _uErrorIdInt := 16#0000_0000;       // 故障码清零（Fault code cleared）
    IF (_ePhase = E_DL_MixPhase.eFault) OR (_ePhase = E_DL_MixPhase.eAbort)
    OR (_ePhase = E_DL_MixPhase.eDone) OR (_ePhase = E_DL_MixPhase.eNg) THEN
        _ePhase := E_DL_MixPhase.eIdle; // 故障/中止/完成/不合格态回空闲（Terminal phases back to idle）
        _bRunIssued := FALSE;           // 运行锁存撤销（Run latch revoked）
        _bConfirmed := FALSE;
        _bRevPending := FALSE;
        _bRevInStop := FALSE;
        _tElapsedInt := T#0S;           // 计时清零（Elapsed reset）
    END_IF
END_IF

// ============================================================================
// 段 3｜中止电平与扭矩保护全局监视（优先级最高）
//      Abort level and torque protection global monitors (highest priority)
// ============================================================================
IF bEnable AND (NOT _bFaultLatch) AND (NOT bAbort)
AND ((_ePhase = E_DL_MixPhase.eMixing) OR (_ePhase = E_DL_MixPhase.eVerify)
  OR (_ePhase = E_DL_MixPhase.eDischarge) OR (_ePhase = E_DL_MixPhase.ePreCheck)) THEN
    IF _bFiniteTrq AND (fActTorque >= _fTorqueLimEff) THEN
        _bCmdStopReq := TRUE;           // 扭矩超限立即停（Torque over limit, stop now）
        _bFaultLatch := TRUE;
        _uErrorIdInt := DL_MIX_ERR_TORQUE;   // 0005_0263 扭矩超保护上限（疑似卡桨）【故障级】/ Torque over limit, fault level
        _ePhase := E_DL_MixPhase.eFault;
    END_IF
END_IF

// 中止电平：任意执行相 → 立即停转、禁止出料、判定作废（Abort level intercept）
IF bEnable AND bAbort AND (NOT _bFaultLatch)
AND (_ePhase <> E_DL_MixPhase.eIdle) AND (_ePhase <> E_DL_MixPhase.eFault)
AND (_ePhase <> E_DL_MixPhase.eAbort) THEN
    _bCmdStopReq := TRUE;               // 立即停转请求（Immediate stop request）
    _bCmdRunReq := FALSE;               // 撤销一切运动请求（Revoke motion requests）
    _bCmdFreqReq := FALSE;
    _bRevPending := FALSE;
    _bRevInStop := FALSE;
    _ePhase := E_DL_MixPhase.eAbort;    // 进入中止保持态（Enter abort hold）
END_IF

// ============================================================================
// 段 4｜核心相位状态机（ENUM + CASE，含 ELSE 非法状态兜底）
//      Core phase state machine (ENUM + CASE with ELSE fallback)
// ============================================================================
IF bEnable AND (NOT _bFaultLatch) AND (NOT bAbort) THEN
    CASE _ePhase OF

        E_DL_MixPhase.eIdle: // 空闲：等启动沿
            IF _fbTrigStart.Q AND (NOT iDrive.bFault) THEN
                _ePhase := E_DL_MixPhase.ePreCheck;      // 受理启动（Start accepted）
                _tElapsedInt := T#0S;                    // 计时清零（Elapsed reset）
                tElapsed := T#0S;                        // 出口计时清零（Outlet elapsed reset）
                _bConfirmed := FALSE;
                _bRunFwd := TRUE;                        // 初始方向正转（Initial direction forward）
                _bDirFwd := TRUE;
            END_IF

        E_DL_MixPhase.ePreCheck: // 前置确认：料已投 + 出料阀关 + 驱动无故障（偏离留档①判据）
            IF bMaterialReady AND bOutletClosed AND (NOT iDrive.bFault) THEN
                _bConfirmed := FALSE;                    // 确认标志复位（Confirm flag reset）
                _fFreqLast := 0.0;                       // 末次下发频率清零（Last sent reset）
                _bCmdFreqReq := TRUE;                    // 登记频率设定（Register setpoint）
                _fFreqReq := _fSetEff;
                _bCmdRunReq := TRUE;                     // 调度器 Run 优先：本拍发运行，设定下一拍补发（Run dispatches first, setpoint follows）
                _bRunFwd := _bDirFwd;
                _ePhase := E_DL_MixPhase.eMixing;        // 进入搅拌（Enter mixing）
            ELSIF _fbTonPreChk.Q THEN
                _bFaultLatch := TRUE;                    // 前置确认超时（Precheck timeout）
                _uErrorIdInt := DL_MIX_ERR_PRECHK;       // 0005_0260 前置条件不成立【故障级】/ Precheck failed, fault level
                _ePhase := E_DL_MixPhase.eFault;
            END_IF

        E_DL_MixPhase.eMixing: // 搅拌：确认窗监视 + 计时 + 交替换向 + 终点判据
            IF (NOT _bConfirmed) AND _bFiniteSpd
            AND (fActSpeed >= _fSetEff * DL_MIX_SPD_OK_FRAC) THEN
                _bConfirmed := TRUE;                     // 转速确认通过（Speed confirmed）
            END_IF
            IF _fbTonSpdChk.Q AND (NOT _bConfirmed) THEN
                _bCmdStopReq := TRUE;                    // 确认失败停机（Stop on confirm failure）
                _bFaultLatch := TRUE;
                _uErrorIdInt := DL_MIX_ERR_SPEED;        // 0005_0261 转速未建立【故障级】/ Speed not established, fault level
                _ePhase := E_DL_MixPhase.eFault;
            ELSE
                IF _bRunIssued AND (NOT _bCmdStopReq) AND (NOT _bCmdRunReq) THEN
                    _bConfirmed := _bConfirmed AND (NOT _bRevInStop); // 停转步期间冻结确认态（Confirm frozen in stop step）
                END_IF
                IF _bConfirmed THEN
                    _tElapsedInt := _tElapsedInt + tCycle;   // 计时仅确认后累计（Elapsed accumulates after confirm）
                    tElapsed := _tElapsedInt;                // 出口计时同步（Outlet elapsed sync）
                END_IF
                // 交替换向三步序：交替周期到 → 登记换向（Alt period reached: arm reversal）
                IF _fbTonAlt.Q THEN
                    _bRevPending := TRUE;                // 换向请求登记（Reversal armed）
                END_IF
                IF _bRevPending AND (NOT _bRevInStop) THEN
                    _bRevInStop := TRUE;                 // 第一步：停转（Step 1: stop）
                    _bCmdStopReq := TRUE;
                END_IF
                IF _bRevInStop AND _bFiniteSpd AND (fActSpeed < DL_MIX_STOP_EPS) THEN
                    // 第二步：转速落零后换向再启（Step 2: restart reversed after standstill）
                    _bDirFwd := NOT _bDirFwd;            // 方向翻转（Direction toggled）
                    _bRunFwd := _bDirFwd;
                    _bCmdRunReq := TRUE;                 // 先发运行（Run first）
                    _fFreqReq := _fSetEff;               // 下一拍补发设定（Frequency follows next scan）
                    _bCmdFreqReq := TRUE;
                    _bRevPending := FALSE;               // 换向序列结束（Reversal sequence done）
                    _bRevInStop := FALSE;
                END_IF
                // 设定变化超容差补发（Resend setpoint beyond epsilon）
                IF _bConfirmed AND (NOT _bRevPending) AND (NOT _bRevInStop)
                AND (ABS(_fSetEff - _fFreqLast) > DL_MIX_FREQ_EPS) THEN
                    _fFreqReq := _fSetEff;               // 登记新设定（Register new setpoint）
                    _bCmdFreqReq := TRUE;
                END_IF
                // 终点判据（End criteria）：已达终点者优先，其次最长超时判 NG
                // 顺序不可倒置：tMixEff ≤ tMixMaxEff 恒成立（段 2 对调自修复），
                // 若「时间终点」排在「最长超时」之后，则 eNg 被完全遮蔽、终态
                // 不可达；此处显式区分终点类型，兼得可达性与时间模式无回归。
                IF bEndByTorque AND _bFiniteTrq AND (fActTorque >= _fTorqueTgtEff) THEN
                    _uInfoCode := DL_MIX_INFO_TORQEND;   // 0005_0163 扭矩终点触发【信息级】/ Torque end reached, info level
                    _ePhase := E_DL_MixPhase.eVerify;    // 进入终点确认（Enter verify）
                ELSIF (NOT bEndByTorque) AND (_tElapsedInt >= _tMixEff) THEN
                    _ePhase := E_DL_MixPhase.eVerify;    // 时间终点（Time end）
                ELSIF _tElapsedInt >= _tMixMaxEff THEN
                    _uInfoCode := DL_MIX_INFO_MAXT;      // 0005_0162 最长混合时间到【信息级】/ Max time reached, info level
                    _bCmdStopReq := TRUE;                // 判 NG 停机（Stop on NG）
                    bNg := TRUE;                         // 不合格出口（NG outlet）
                    bDone := TRUE;                       // 完成单拍（R25 本拍闭环）/ Done pulse (R25)
                    _ePhase := E_DL_MixPhase.eNg;
                END_IF
            END_IF

        E_DL_MixPhase.eVerify: // 终点确认：稳速容差内确认后锁存进料
            IF _bFiniteSpd AND (ABS(fActSpeed - _fSetEff) <= _fSetEff * DL_MIX_VERIFY_FRAC) THEN
                _fFreqReq := DL_MIX_DISCHARGE_SPD;       // 出料助排慢速设定（Discharge assist setpoint）
                _bCmdFreqReq := TRUE;                    // 登记设定（Register setpoint）
                _ePhase := E_DL_MixPhase.eDischarge;     // 进入出料（Enter discharge）
            END_IF

        E_DL_MixPhase.eDischarge: // 出料中：慢速助排，等出料完成
            IF bDischargeDone THEN
                _bCmdStopReq := TRUE;                    // 出料完成停转（Stop after discharge）
                _ePhase := E_DL_MixPhase.eSpinDown;      // 进入停转（Enter spin-down）
            ELSIF _fbTonDischTo.Q THEN
                _bCmdStopReq := TRUE;                    // 超时停机（Stop on timeout）
                _bFaultLatch := TRUE;
                _uErrorIdInt := DL_MIX_ERR_DISCH;        // 0005_0262 出料超时【故障级】/ Discharge timeout, fault level
                _ePhase := E_DL_MixPhase.eFault;
            END_IF

        E_DL_MixPhase.eSpinDown: // 停转：等待转速落零
            IF _bFiniteSpd AND (fActSpeed < DL_MIX_STOP_EPS) THEN
                bOk := TRUE;                             // 合格出口（OK outlet）
                bDone := TRUE;                           // 完成单拍（R25 本拍闭环）/ Done pulse (R25)
                _ePhase := E_DL_MixPhase.eDone;          // 进入完成保持（Enter done hold）
            END_IF

        E_DL_MixPhase.eDone: // 完成保持：判定每拍重算保持（复位路径在段 2）
            bOk := TRUE;                             // 合格保持（OK verdict held every scan）

        E_DL_MixPhase.eNg: // 不合格保持：判定每拍重算保持
            bNg := TRUE;                             // 不合格保持（NG verdict held every scan）

        E_DL_MixPhase.eAbort: // 中止保持：停转完成，禁止出料，等复位
            // 等复位（Awaiting reset）

        E_DL_MixPhase.eFault: // 故障锁存：等复位
            // 等复位（Awaiting reset）

        ELSE // 非法状态兜底（本块专用码位）
            _bCmdStopReq := TRUE;               // 非法状态立即停（Stop on illegal state）
            _bFaultLatch := TRUE;
            _uErrorIdInt := DL_MIX_ERR_STATE;   // 0005_0265 非法状态兜底【故障级】/ Illegal state fallback, fault level
            _ePhase := E_DL_MixPhase.eFault;
    END_CASE
END_IF

// ============================================================================
// 段 5｜接口单发指令调度器（公约 0.13：每拍至多一次方法调用，结构保证）
//      Interface single-shot dispatcher (0.13: at most one method call per scan)
// ============================================================================
IF NOT bEnable THEN
    _bCmdRunReq := FALSE;               // 使能撤销撤销全部请求（Disable revokes all requests）
    _bCmdFreqReq := FALSE;
    _bRunIssued := FALSE;               // 运行锁存撤销（Run latch revoked）
    IF _ePhase <> E_DL_MixPhase.eIdle THEN
        _bCmdStopReq := TRUE;           // 残余运行先停（Stop residual run）
    END_IF
END_IF

IF _bCmdStopReq THEN
    IF iDrive.CmdStop() THEN            // 停止指令无条件受理（Stop unconditionally accepted）
        _bCmdStopReq := FALSE;          // 消费请求（Consume request）
        _bCmdRunReq := FALSE;           // 停止优先：清运行/设定请求（Stop clears run/freq requests）
        _bCmdFreqReq := FALSE;
        _bRunIssued := FALSE;           // 运行锁存撤销（Run latch revoked）
        _fFreqLast := 0.0;              // 末次设定清零（Last setpoint reset）
    END_IF
ELSIF _bCmdRunReq THEN
    IF iDrive.CmdRun(bFwd := _bRunFwd) THEN   // 运行指令（Run command with direction）
        _bCmdRunReq := FALSE;           // 消费请求（Consume request）
        _bRunIssued := TRUE;            // 运行锁存登记（Run latch registered）
    END_IF
ELSIF _bCmdFreqReq THEN
    IF iDrive.SetFrequency(fHz := _fFreqReq) THEN   // 设定指令（SetFrequency command）
        _bCmdFreqReq := FALSE;          // 消费请求（Consume request）
        _fFreqLast := _fFreqReq;        // 登记末次下发（Register last sent）
    END_IF
END_IF

// ============================================================================
// 段 6｜出口派生（方向互斥断言由同源派生保证；进度折算除前判零）
//      Outlet derivation (mutual exclusion by common source; progress divide guarded)
// ============================================================================
bDirForward := _bRunIssued AND _bDirFwd;             // 正转出口（Forward outlet）
bDirReverse := _bRunIssued AND (NOT _bDirFwd);       // 反转出口（Reverse outlet），与正转同源互斥 / Mutually exclusive by source

IF (_ePhase = E_DL_MixPhase.eDischarge) AND _bRunIssued THEN
    fSpeedCmd := DL_MIX_DISCHARGE_SPD;               // 出料助排慢速（Discharge assist speed）
ELSIF _bRunIssued THEN
    fSpeedCmd := _fSetEff;                           // 搅拌设定转速（Mixing setpoint）
ELSE
    fSpeedCmd := 0.0;                                // 停转（Standstill）
END_IF

// 进度折算：已混合秒值/目标秒值 [-]，钳位 [0,1]（R20 量纲：无量纲）
// Progress: elapsed seconds / target seconds, clamped 0..1 (dimensionless per R20)
IF TIME_TO_REAL(_tMixEff) > DL_MIX_EPS THEN
    fProgress := LIMIT(0.0, TIME_TO_REAL(_tElapsedInt) / TIME_TO_REAL(_tMixEff), 1.0);
END_IF

// 判定互斥出口断言（规格 §6-8）：OK 与 NG 恒不同真，冲突时 NG 优先
// Verdict mutual-exclusion assertion: OK and NG never both TRUE, NG wins
IF bOk AND bNg THEN
    bOk := FALSE;                                    // 不合格优先（NG priority）
END_IF

bBusy := (_ePhase = E_DL_MixPhase.ePreCheck)
      OR (_ePhase = E_DL_MixPhase.eMixing)
      OR (_ePhase = E_DL_MixPhase.eVerify)
      OR (_ePhase = E_DL_MixPhase.eDischarge)
      OR (_ePhase = E_DL_MixPhase.eSpinDown);        // 执行中派生（Busy derived）

ePhase := _ePhase;                       // 相位镜像（Phase mirror）

// ============================================================================
// 段 7｜bError/uErrorId 出口（R21：bError 显式排除信息级码）
//      Outlets: bError excludes info codes (R21)
// ============================================================================
bError := _bFaultLatch;                  // 故障级派生式（Fault-level derived form）
IF _bFaultLatch THEN
    uErrorId := _uErrorIdInt;            // 故障级码优先透出（Fault-level priority）
ELSE
    uErrorId := _uInfoCode;              // 无故障时透出本拍信息级码（Transient info code）
END_IF
END_FUNCTION_BLOCK
